(* Asserts that parse rejects header with the expected reason and allocates nothing. *)
METHOD _expectRejected
VAR_INPUT
	header: T_MaxString;
	expected: E_TraceStateFailureReason;
END_VAR
VAR
	_pTraceState: POINTER TO FB_TraceState;
	_success: BOOL;
	_reason: E_TraceStateFailureReason;
END_VAR
_success := TraceStateFactory.parse(pDest:=_pTraceState, pHeader:=ADR(header), failureReason=>_reason);
THIS^.AssertFalse(_success, CONCAT('Expected parse to reject: ', header));
THIS^.AssertEquals_UDINT(TO_UDINT(expected), TO_UDINT(_reason), CONCAT('Expected the failure reason for: ', header));
THIS^.AssertTrue(_pTraceState = 0, CONCAT('Expected nothing to be allocated for: ', header));
IF _pTraceState <> 0 THEN _pTraceState^.delete(pSelf:=_pTraceState); END_IF
END_METHOD

(*
	Writes a valid 515 character header: four 128 character entries k0..k3 joined by ','.
	It is built byte by byte because STRING functions stop at 255 characters.
*)
METHOD _fillLongHeader
VAR_IN_OUT
	header: STRING(600);
END_VAR
VAR
	_p: POINTER TO BYTE;
	_entry: UDINT;
	_i: UDINT;
	_n: UDINT;
END_VAR
_p := ADR(header);
FOR _entry := 0 TO 3 DO
	IF _entry > 0 THEN
		_p[_n] := 16#2C;  // ','
		_n := _n + 1;
	END_IF
	_p[_n] := 16#6B;  // 'k'
	_p[_n + 1] := 16#30 + TO_BYTE(_entry);
	_p[_n + 2] := 16#3D;  // '='
	_n := _n + 3;
	FOR _i := 1 TO 125 DO
		_p[_n] := 16#61 + TO_BYTE(_i MOD 26);
		_n := _n + 1;
	END_FOR
END_FOR
_p[_n] := 0;
END_METHOD

(* parse drops empty members and the optional whitespace around ',' and keeps the order. *)
METHOD testParseCanonicalises : REFERENCE TO FB_Test
VAR
	header: T_MaxString := ' vendor=abc ,, rojo=00f067aa0ba902b7$T, congo@t61rcwkgmze=x ';
	expected: T_MaxString := 'vendor=abc,rojo=00f067aa0ba902b7,congo@t61rcwkgmze=x';
	pTraceState: POINTER TO FB_TraceState;
	success: BOOL;
	reason: E_TraceStateFailureReason;
END_VAR
TcUnit.TEST('testParseCanonicalises');
	success := TraceStateFactory.parse(pDest:=pTraceState, pHeader:=ADR(header), failureReason=>reason);
	THIS^.AssertTrue(success, 'Expected a valid header to parse');
	THIS^.AssertEquals_UDINT(TO_UDINT(E_TraceStateFailureReason.NA), TO_UDINT(reason), 'Expected no failure reason');
	THIS^.AssertTrue(pTraceState <> 0, 'Expected a trace state');
	IF pTraceState <> 0 THEN
		THIS^.AssertEquals_STRING(expected, pTraceState^.pString^, 'Expected the canonical header');
		THIS^.AssertEquals_UDINT(TO_UDINT(LEN(expected)), pTraceState^.length, 'Expected the canonical length');
		THIS^.AssertEquals_UDINT(3, pTraceState^.count, 'Expected three entries');
		pTraceState^.delete(pSelf:=pTraceState);
		THIS^.AssertTrue(pTraceState = 0, 'Expected delete to clear the pointer');
	END_IF
TcUnit.TEST_FINISHED();
END_METHOD

(* An empty header, or one of only empty members, is valid but holds nothing, so no trace state is allocated. *)
METHOD testParseEmptyHeader : REFERENCE TO FB_Test
VAR
	empty: T_MaxString := '';
	blank: T_MaxString := ' , ,,$T';
	pTraceState: POINTER TO FB_TraceState;
	success: BOOL;
	reason: E_TraceStateFailureReason;
END_VAR
TcUnit.TEST('testParseEmptyHeader');
	success := TraceStateFactory.parse(pDest:=pTraceState, pHeader:=ADR(empty), failureReason=>reason);
	THIS^.AssertTrue(success, 'Expected an empty header to be accepted');
	THIS^.AssertEquals_UDINT(TO_UDINT(E_TraceStateFailureReason.NA), TO_UDINT(reason), 'Expected no failure reason');
	THIS^.AssertTrue(pTraceState = 0, 'Expected no trace state for an empty header');

	success := TraceStateFactory.parse(pDest:=pTraceState, pHeader:=ADR(blank), failureReason=>reason);
	THIS^.AssertTrue(success, 'Expected a header of empty members to be accepted');
	THIS^.AssertTrue(pTraceState = 0, 'Expected no trace state for a header of empty members');
	IF pTraceState <> 0 THEN pTraceState^.delete(pSelf:=pTraceState); END_IF
TcUnit.TEST_FINISHED();
END_METHOD

(* Anything that breaks the W3C key or value grammar, or repeats a key, is rejected whole. *)
METHOD testParseRejectsInvalidHeaders : REFERENCE TO FB_Test
VAR
	pTraceState: POINTER TO FB_TraceState;
	pOther: POINTER TO FB_TraceState;
	header: T_MaxString := 'vendor=abc';
	success: BOOL;
	reason: E_TraceStateFailureReason;
END_VAR
TcUnit.TEST('testParseRejectsInvalidHeaders');
	THIS^._expectRejected(header:='Vendor=abc', expected:=E_TraceStateFailureReason.INVALID_KEY);
	THIS^._expectRejected(header:='1vendor=x', expected:=E_TraceStateFailureReason.INVALID_KEY);
	THIS^._expectRejected(header:='=x', expected:=E_TraceStateFailureReason.INVALID_KEY);
	THIS^._expectRejected(header:='@sys=x', expected:=E_TraceStateFailureReason.INVALID_KEY);
	THIS^._expectRejected(header:='tenant@=x', expected:=E_TraceStateFailureReason.INVALID_KEY);
	THIS^._expectRejected(header:='tenant@1sys=x', expected:=E_TraceStateFailureReason.INVALID_KEY);
	THIS^._expectRejected(header:='a@b@c=x', expected:=E_TraceStateFailureReason.INVALID_KEY);
	THIS^._expectRejected(header:='ven dor=x', expected:=E_TraceStateFailureReason.INVALID_KEY);
	THIS^._expectRejected(header:='vendor', expected:=E_TraceStateFailureReason.INVALID_VALUE);
	THIS^._expectRejected(header:='vendor=', expected:=E_TraceStateFailureReason.INVALID_VALUE);
	THIS^._expectRejected(header:='vendor=a=b', expected:=E_TraceStateFailureReason.INVALID_VALUE);
	THIS^._expectRejected(header:='vendor=a$Tb', expected:=E_TraceStateFailureReason.INVALID_VALUE);
	THIS^._expectRejected(header:='good=1,vendor=a=b', expected:=E_TraceStateFailureReason.INVALID_VALUE);
	THIS^._expectRejected(header:='a=1,b=2,a=3', expected:=E_TraceStateFailureReason.DUPLICATE_KEY);

	success := TraceStateFactory.parse(pDest:=pTraceState, pHeader:=0, failureReason=>reason);
	THIS^.AssertFalse(success, 'Expected a null header pointer to be rejected');
	THIS^.AssertEquals_UDINT(TO_UDINT(E_TraceStateFailureReason.HEADER_POINTER_NULL), TO_UDINT(reason), 'Expected HEADER_POINTER_NULL');

	TraceStateFactory.parse(pDest:=pTraceState, pHeader:=ADR(header));
	pOther := pTraceState;
	success := TraceStateFactory.parse(pDest:=pTraceState, pHeader:=ADR(header), failureReason=>reason);
	THIS^.AssertFalse(success, 'Expected an assigned destination to be rejected');
	THIS^.AssertEquals_UDINT(TO_UDINT(E_TraceStateFailureReason.DESTINATION_ALREADY_ASSIGNED), TO_UDINT(reason), 'Expected DESTINATION_ALREADY_ASSIGNED');
	THIS^.AssertTrue(pTraceState = pOther, 'Expected the destination to be left alone');
	IF pTraceState <> 0 THEN pTraceState^.delete(pSelf:=pTraceState); END_IF
TcUnit.TEST_FINISHED();
END_METHOD

(* W3C allows at most 32 entries; a 33rd is rejected. *)
METHOD testParseEntryLimit : REFERENCE TO FB_Test
VAR
	header: T_MaxString;
	i: UDINT;
	pTraceState: POINTER TO FB_TraceState;
	success: BOOL;
	reason: E_TraceStateFailureReason;
END_VAR
TcUnit.TEST('testParseEntryLimit');
	header := 'k0=1';
	FOR i := 1 TO 31 DO
		header := CONCAT(header, CONCAT(CONCAT(',k', UDINT_TO_STRING(i)), '=1'));
	END_FOR
	success := TraceStateFactory.parse(pDest:=pTraceState, pHeader:=ADR(header), failureReason=>reason);
	THIS^.AssertTrue(success, 'Expected 32 entries to be accepted');
	IF pTraceState <> 0 THEN
		THIS^.AssertEquals_UDINT(32, pTraceState^.count, 'Expected 32 entries');
		pTraceState^.delete(pSelf:=pTraceState);
	END_IF

	header := CONCAT(header, ',k32=1');
	success := TraceStateFactory.parse(pDest:=pTraceState, pHeader:=ADR(header), failureReason=>reason);
	THIS^.AssertFalse(success, 'Expected 33 entries to be rejected');
	THIS^.AssertEquals_UDINT(TO_UDINT(E_TraceStateFailureReason.TOO_MANY_ENTRIES), TO_UDINT(reason), 'Expected TOO_MANY_ENTRIES');
	THIS^.AssertTrue(pTraceState = 0, 'Expected nothing to be allocated');
TcUnit.TEST_FINISHED();
END_METHOD

(* A header longer than T_MaxString is kept whole; W3C asks for at least 512 characters. *)
METHOD testParseLongHeader : REFERENCE TO FB_Test
VAR
	header: STRING(600);
	pTraceState: POINTER TO FB_TraceState;
	success: BOOL;
END_VAR
TcUnit.TEST('testParseLongHeader');
	THIS^._fillLongHeader(header:=header);
	THIS^.AssertEquals_UDINT(515, TO_UDINT(LEN2(ADR(header))), 'Expected a 515 character test header');
	success := TraceStateFactory.parse(pDest:=pTraceState, pHeader:=ADR(header));
	THIS^.AssertTrue(success, 'Expected the long header to parse');
	IF pTraceState <> 0 THEN
		THIS^.AssertEquals_UDINT(515, pTraceState^.length, 'Expected all 515 characters');
		THIS^.AssertEquals_UDINT(4, pTraceState^.count, 'Expected four entries');
		THIS^.AssertTrue(MEMCMP(pTraceState^.pString, ADR(header), 516) = 0, 'Expected the header unchanged, with its terminator');
		pTraceState^.delete(pSelf:=pTraceState);
	END_IF
TcUnit.TEST_FINISHED();
END_METHOD

(* clone owns its own buffer, so it outlives the source. *)
METHOD testCloneIsIndependent : REFERENCE TO FB_Test
VAR
	header: T_MaxString := 'vendor=abc,rojo=1';
	pSource: POINTER TO FB_TraceState;
	pClone: POINTER TO FB_TraceState;
	pOther: POINTER TO FB_TraceState;
	success: BOOL;
	reason: E_TraceStateFailureReason;
END_VAR
TcUnit.TEST('testCloneIsIndependent');
	TraceStateFactory.parse(pDest:=pSource, pHeader:=ADR(header));
	success := TraceStateFactory.clone(pDest:=pClone, pSrc:=pSource, failureReason=>reason);
	THIS^.AssertTrue(success, 'Expected clone to succeed');
	THIS^.AssertTrue(pClone <> 0 AND pClone <> pSource, 'Expected a new trace state');
	IF pSource <> 0 AND pClone <> 0 THEN
		THIS^.AssertTrue(pClone^.pString <> pSource^.pString, 'Expected the clone to own its own buffer');
	END_IF

	success := TraceStateFactory.clone(pDest:=pClone, pSrc:=pSource, failureReason=>reason);
	THIS^.AssertFalse(success, 'Expected clone into an assigned destination to fail');
	THIS^.AssertEquals_UDINT(TO_UDINT(E_TraceStateFailureReason.DESTINATION_ALREADY_ASSIGNED), TO_UDINT(reason), 'Expected DESTINATION_ALREADY_ASSIGNED');
	success := TraceStateFactory.clone(pDest:=pOther, pSrc:=0, failureReason=>reason);
	THIS^.AssertFalse(success, 'Expected clone of a null source to fail');
	THIS^.AssertEquals_UDINT(TO_UDINT(E_TraceStateFailureReason.SOURCE_POINTER_NULL), TO_UDINT(reason), 'Expected SOURCE_POINTER_NULL');

	IF pSource <> 0 THEN pSource^.delete(pSelf:=pSource); END_IF
	IF pClone <> 0 THEN
		THIS^.AssertEquals_STRING('vendor=abc,rojo=1', pClone^.pString^, 'Expected the clone to outlive its source');
		THIS^.AssertEquals_UDINT(2, pClone^.count, 'Expected the entry count to be copied');
		pClone^.delete(pSelf:=pClone);
	END_IF
TcUnit.TEST_FINISHED();
END_METHOD

(* truncate removes entries over 128 characters first, then entries from the right, and never cuts an entry. *)
METHOD testTruncateFollowsW3C : REFERENCE TO FB_Test
VAR
	header: STRING(600);
	pBytes: POINTER TO BYTE;
	i: UDINT;
	pSource: POINTER TO FB_TraceState;
	pResult: POINTER TO FB_TraceState;
	success: BOOL;
	reason: E_TraceStateFailureReason;
END_VAR
TcUnit.TEST('testTruncateFollowsW3C');
	// a=1,big=<130 characters>,b=2,c=3
	header := 'a=1,big=';
	pBytes := ADR(header);
	FOR i := 8 TO 137 DO
		pBytes[i] := 16#78;  // 'x'
	END_FOR
	pBytes[138] := 0;
	MEMCPY(pBytes + 138, ADR(',b=2,c=3'), 9);
	success := TraceStateFactory.parse(pDest:=pSource, pHeader:=ADR(header));
	THIS^.AssertTrue(success AND pSource <> 0, 'Expected the header to parse');
	IF pSource = 0 THEN
		TcUnit.TEST_FINISHED();
		RETURN;
	END_IF
	THIS^.AssertEquals_UDINT(146, pSource^.length, 'Expected a 146 character test header');

	success := TraceStateFactory.truncate(pDest:=pResult, pSrc:=pSource, maxLength:=1000, failureReason=>reason);
	THIS^.AssertTrue(success AND pResult <> 0, 'Expected a header that fits to be copied');
	IF pResult <> 0 THEN
		THIS^.AssertTrue(pResult <> pSource AND pResult^.length = 146, 'Expected a whole copy');
		pResult^.delete(pSelf:=pResult);
	END_IF

	success := TraceStateFactory.truncate(pDest:=pResult, pSrc:=pSource, maxLength:=20, failureReason=>reason);
	THIS^.AssertTrue(success, 'Expected truncate to succeed');
	IF pResult <> 0 THEN
		THIS^.AssertEquals_STRING('a=1,b=2,c=3', pResult^.pString^, 'Expected the large entry to go first');
		THIS^.AssertEquals_UDINT(3, pResult^.count, 'Expected three entries');
		pResult^.delete(pSelf:=pResult);
	ELSE
		THIS^.AssertTrue(FALSE, 'Expected a truncated trace state');
	END_IF

	success := TraceStateFactory.truncate(pDest:=pResult, pSrc:=pSource, maxLength:=7, failureReason=>reason);
	THIS^.AssertTrue(success, 'Expected truncate to succeed');
	IF pResult <> 0 THEN
		THIS^.AssertEquals_STRING('a=1,b=2', pResult^.pString^, 'Expected entries to go from the right next');
		pResult^.delete(pSelf:=pResult);
	ELSE
		THIS^.AssertTrue(FALSE, 'Expected a truncated trace state');
	END_IF

	success := TraceStateFactory.truncate(pDest:=pResult, pSrc:=pSource, maxLength:=2, failureReason=>reason);
	THIS^.AssertTrue(success, 'Expected truncate to succeed when nothing fits');
	THIS^.AssertTrue(pResult = 0, 'Expected no trace state when no entry fits');
	IF pResult <> 0 THEN pResult^.delete(pSelf:=pResult); END_IF

	success := TraceStateFactory.truncate(pDest:=pResult, pSrc:=0, maxLength:=512, failureReason=>reason);
	THIS^.AssertFalse(success, 'Expected a null source to be rejected');
	THIS^.AssertEquals_UDINT(TO_UDINT(E_TraceStateFailureReason.SOURCE_POINTER_NULL), TO_UDINT(reason), 'Expected SOURCE_POINTER_NULL');

	pSource^.delete(pSelf:=pSource);
TcUnit.TEST_FINISHED();
END_METHOD

END_FUNCTION_BLOCK

// ---- TEST/TRACING/PROPAGATION/FB_TestTraceContextPropagator.TcPOU
(* Tests TraceContextPropagator.extract and inject against the W3C traceparent and tracestate rules. *)
FUNCTION_BLOCK FB_TestTraceContextPropagator EXTENDS FB_TestSuite

THIS^.testExtractsTraceparentAndTracestate();
THIS^.testKeepsUnsampledFlag();
THIS^.testAcceptsFutureVersion();
THIS^.testMeasuresTraceparentBeyond255();
THIS^.testTracestateIsOptional();
THIS^.testKeepsLongTracestateWhole();
THIS^.testRejectsMalformedTraceparent();
THIS^.testRejectsAssignedDestination();
THIS^.testInjectWritesExtractedCarrier();
THIS^.testInjectDropsWholeTracestateEntries();
THIS^.testInjectRejectsMissingOrInvalidContext();

(*
	Asserts that extract rejects traceparent with the expected reason and leaves the destination
	at 0. The tracestate beside it is valid, so this also shows a bad traceparent drops it.
*)
METHOD _expectRejected
VAR_INPUT
	traceparent: T_MaxString;  // longer than 55, so overlong headers reach extract whole
	expected: E_PropagationFailureReason;
END_VAR
VAR
	_pContext: POINTER TO FB_SpanContext;
	_success: BOOL;
	_reason: E_PropagationFailureReason;
END_VAR
_success := TraceContextPropagator.extract(
	pDest:=_pContext,
	traceparent:=traceparent,
	tracestate:='vendor=abc',
	failureReason=>_reason
);
THIS^.AssertFalse(_success, CONCAT('Expected extract to reject: ', traceparent));
THIS^.AssertEquals_UDINT(TO_UDINT(expected), TO_UDINT(_reason), CONCAT('Expected the failure reason for: ', traceparent));
THIS^.AssertTrue(_pContext = 0, CONCAT('Expected no context for: ', traceparent));
IF _pContext <> 0 THEN _pContext^.delete(pSelf:=_pContext); END_IF
END_METHOD

(*
	The W3C example carrier becomes a remote context holding the caller's trace id, span id,
	sampled bit and tracestate, so a PLC span can link back to the span that triggered it.
*)
METHOD testExtractsTraceparentAndTracestate : REFERENCE TO FB_Test
VAR
	traceparent: STRING(55) := '00-4bf92f3577b34da6a3ce929d0e0e4736-00f067aa0ba902b7-01';
	tracestate: STRING(512) := 'congo=t61rcWkgMzE,rojo=00f067aa0ba902b7';
	expectedTraceId: ARRAY [0..15] OF BYTE := [
		16#4B, 16#F9, 16#2F, 16#35, 16#77, 16#B3, 16#4D, 16#A6,
		16#A3, 16#CE, 16#92, 16#9D, 16#0E, 16#0E, 16#47, 16#36];
	expectedSpanId: ARRAY [0..7] OF BYTE := [16#00, 16#F0, 16#67, 16#AA, 16#0B, 16#A9, 16#02, 16#B7];
	pContext: POINTER TO FB_SpanContext;
	pTraceState: POINTER TO FB_TraceState;
	traceId: REFERENCE TO FB_TraceId;
	spanId: REFERENCE TO FB_SpanId;
	success: BOOL;
	reason: E_PropagationFailureReason;
END_VAR
TcUnit.TEST('testExtractsTraceparentAndTracestate');
	success := TraceContextPropagator.extract(
		pDest:=pContext,
		traceparent:=traceparent,
		tracestate:=tracestate,
		failureReason=>reason
	);
	THIS^.AssertTrue(success, 'Expected the W3C example carrier to be extracted');
	THIS^.AssertEquals_UDINT(TO_UDINT(E_PropagationFailureReason.NA), TO_UDINT(reason), 'Expected no failure reason on success');
	THIS^.AssertTrue(pContext <> 0, 'Expected extract to assign the destination');
	IF pContext = 0 THEN
		TcUnit.TEST_FINISHED();
		RETURN;
	END_IF

	traceId REF= pContext^.traceId;
	spanId REF= pContext^.spanId;
	THIS^.AssertTrue(
		MEMCMP(ADR(traceId.bytes), ADR(expectedTraceId), SIZEOF(expectedTraceId)) = 0,
		'Expected the trace id decoded from the traceparent'
	);
	THIS^.AssertTrue(
		MEMCMP(ADR(spanId.bytes), ADR(expectedSpanId), SIZEOF(expectedSpanId)) = 0,
		'Expected the caller$'s span id decoded from the traceparent'
	);
	THIS^.AssertEquals_UDINT(16#301, pContext^.traceFlags, 'Expected the sampled bit and both remote bits');
	THIS^.AssertTrue(pContext^.isRemote(), 'Expected an extracted context to be remote');

	pTraceState := pContext^.traceState;
	THIS^.AssertTrue(pTraceState <> 0, 'Expected the tracestate to be kept');
	IF pTraceState <> 0 THEN
		THIS^.AssertEquals_STRING('congo=t61rcWkgMzE,rojo=00f067aa0ba902b7', pTraceState^.pString^, 'Expected the tracestate entries in their original order');
	END_IF
	pContext^.delete(pSelf:=pContext);
TcUnit.TEST_FINISHED();
END_METHOD

(*
	A caller that did not sample its own trace still produces a context: the sampled bit is
	carried as sent, and the default sampler does not sample a child of the context.
*)
METHOD testKeepsUnsampledFlag : REFERENCE TO FB_Test
VAR
	traceparent: STRING(55) := '00-4bf92f3577b34da6a3ce929d0e0e4736-00f067aa0ba902b7-00';
	pContext: POINTER TO FB_SpanContext;
	success: BOOL;
END_VAR
TcUnit.TEST('testKeepsUnsampledFlag');
	success := TraceContextPropagator.extract(pDest:=pContext, traceparent:=traceparent, tracestate:='');
	THIS^.AssertTrue(success, 'Expected an unsampled carrier to be extracted');
	IF pContext <> 0 THEN
		THIS^.AssertEquals_UDINT(16#300, pContext^.traceFlags, 'Expected both remote bits and no sampled bit');
		THIS^.AssertTrue(pContext^.isRemote(), 'Expected an extracted context to be remote');
		pContext^.delete(pSelf:=pContext);
	END_IF
TcUnit.TEST_FINISHED();
END_METHOD

(*
	W3C asks a parser to read a newer version as version 00 rather than reject it, ignoring any
	fields after the flags, so a caller that upgrades its tracing library does not lose the link.
	The flags may end the header or be followed by '-' and more fields.
*)
METHOD testAcceptsFutureVersion : REFERENCE TO FB_Test
VAR
	traceparent: STRING(80) := 'cc-4bf92f3577b34da6a3ce929d0e0e4736-00f067aa0ba902b7-01-newfield';
	traceparentWithoutFields: STRING(55) := 'cc-4bf92f3577b34da6a3ce929d0e0e4736-00f067aa0ba902b7-01';
	pContext: POINTER TO FB_SpanContext;
	success: BOOL;
	reason: E_PropagationFailureReason;
END_VAR
TcUnit.TEST('testAcceptsFutureVersion');
	success := TraceContextPropagator.extract(pDest:=pContext, traceparent:=traceparent, tracestate:='', failureReason=>reason);
	THIS^.AssertTrue(success, 'Expected version cc with an extra field to be read as version 00');
	THIS^.AssertEquals_UDINT(TO_UDINT(E_PropagationFailureReason.NA), TO_UDINT(reason), 'Expected no failure reason for a future version');
	IF pContext <> 0 THEN pContext^.delete(pSelf:=pContext); END_IF

	// the flags end the header
	success := TraceContextPropagator.extract(pDest:=pContext, traceparent:=traceparentWithoutFields, tracestate:='', failureReason=>reason);
	THIS^.AssertTrue(success, 'Expected version cc with no extra field to be read as version 00');
	THIS^.AssertEquals_UDINT(TO_UDINT(E_PropagationFailureReason.NA), TO_UDINT(reason), 'Expected no failure reason for a 55 character future version');
	IF pContext <> 0 THEN pContext^.delete(pSelf:=pContext); END_IF
TcUnit.TEST_FINISHED();
END_METHOD

(*
	The traceparent alone identifies the caller's span. A missing tracestate, or one that breaks
	the W3C grammar, leaves the context without a trace state instead of failing the extraction.
*)
METHOD testTracestateIsOptional : REFERENCE TO FB_Test
VAR
	traceparent: STRING(55) := '00-4bf92f3577b34da6a3ce929d0e0e4736-00f067aa0ba902b7-01';
	pContext: POINTER TO FB_SpanContext;
	success: BOOL;
	reason: E_PropagationFailureReason;
END_VAR
TcUnit.TEST('testTracestateIsOptional');
	// no tracestate header
	success := TraceContextPropagator.extract(pDest:=pContext, traceparent:=traceparent, tracestate:='', failureReason=>reason);
	THIS^.AssertTrue(success, 'Expected a carrier without tracestate to be extracted');
	THIS^.AssertTrue(pContext <> 0 AND_THEN pContext^.traceState = 0, 'Expected no trace state without a tracestate header');
	IF pContext <> 0 THEN pContext^.delete(pSelf:=pContext); END_IF

	// an uppercase key breaks the tracestate grammar, so only the trace state is dropped
	success := TraceContextPropagator.extract(pDest:=pContext, traceparent:=traceparent, tracestate:='Vendor=abc', failureReason=>reason);
	THIS^.AssertTrue(success, 'Expected an invalid tracestate not to fail the extraction');
	THIS^.AssertEquals_UDINT(TO_UDINT(E_PropagationFailureReason.NA), TO_UDINT(reason), 'Expected no failure reason for a dropped tracestate');
	THIS^.AssertTrue(pContext <> 0 AND_THEN pContext^.traceState = 0, 'Expected an invalid tracestate to be dropped');
	IF pContext <> 0 THEN pContext^.delete(pSelf:=pContext); END_IF
TcUnit.TEST_FINISHED();
END_METHOD

(*
	Each way a traceparent can break the W3C format is reported by its own reason, and nothing
	is allocated, so the caller can start an unlinked span and log why.
*)
METHOD testRejectsMalformedTraceparent : REFERENCE TO FB_Test
TcUnit.TEST('testRejectsMalformedTraceparent');
	// no header at all
	THIS^._expectRejected(traceparent:='', expected:=E_PropagationFailureReason.TRACEPARENT_EMPTY);
	// the flags are missing
	THIS^._expectRejected(traceparent:='00-4bf92f3577b34da6a3ce929d0e0e4736-00f067aa0ba902b7', expected:=E_PropagationFailureReason.TRACEPARENT_LENGTH_INVALID);
	// version ff is reserved as invalid
	THIS^._expectRejected(traceparent:='ff-4bf92f3577b34da6a3ce929d0e0e4736-00f067aa0ba902b7-01', expected:=E_PropagationFailureReason.VERSION_INVALID);
	// the version is not hex
	THIS^._expectRejected(traceparent:='0g-4bf92f3577b34da6a3ce929d0e0e4736-00f067aa0ba902b7-01', expected:=E_PropagationFailureReason.VERSION_INVALID);
	// the version is not followed by '-'
	THIS^._expectRejected(traceparent:='00_4bf92f3577b34da6a3ce929d0e0e4736-00f067aa0ba902b7-01', expected:=E_PropagationFailureReason.DELIMITER_INVALID);
	// W3C allows only lowercase hex
	THIS^._expectRejected(traceparent:='00-4BF92F3577B34DA6A3CE929D0E0E4736-00f067aa0ba902b7-01', expected:=E_PropagationFailureReason.TRACE_ID_INVALID);
	// an all-zero trace id means absent
	THIS^._expectRejected(traceparent:='00-00000000000000000000000000000000-00f067aa0ba902b7-01', expected:=E_PropagationFailureReason.TRACE_ID_INVALID);
	// the span id is not hex
	THIS^._expectRejected(traceparent:='00-4bf92f3577b34da6a3ce929d0e0e4736-00f067aa0ba902bx-01', expected:=E_PropagationFailureReason.SPAN_ID_INVALID);
	// an all-zero span id means absent
	THIS^._expectRejected(traceparent:='00-4bf92f3577b34da6a3ce929d0e0e4736-0000000000000000-01', expected:=E_PropagationFailureReason.SPAN_ID_INVALID);
	// the flags are not hex
	THIS^._expectRejected(traceparent:='00-4bf92f3577b34da6a3ce929d0e0e4736-00f067aa0ba902b7-0z', expected:=E_PropagationFailureReason.TRACE_FLAGS_INVALID);
	// version 00 is exactly 55 characters, so nothing may follow the flags
	THIS^._expectRejected(traceparent:='00-4bf92f3577b34da6a3ce929d0e0e4736-00f067aa0ba902b7-01-00', expected:=E_PropagationFailureReason.TRACEPARENT_LENGTH_INVALID);
	// a future version's flags must be followed by '-' or the end of the header
	THIS^._expectRejected(traceparent:='cc-4bf92f3577b34da6a3ce929d0e0e4736-00f067aa0ba902b7-01x', expected:=E_PropagationFailureReason.DELIMITER_INVALID);
TcUnit.TEST_FINISHED();
END_METHOD

(* extract never overwrites a context the caller already owns, which would leak it. *)
METHOD testRejectsAssignedDestination : REFERENCE TO FB_Test
VAR
	traceparent: STRING(55) := '00-4bf92f3577b34da6a3ce929d0e0e4736-00f067aa0ba902b7-01';
	pContext: POINTER TO FB_SpanContext;
	pFirst: POINTER TO FB_SpanContext;
	success: BOOL;
	reason: E_PropagationFailureReason;
END_VAR
TcUnit.TEST('testRejectsAssignedDestination');
	TraceContextPropagator.extract(pDest:=pContext, traceparent:=traceparent, tracestate:='');
	pFirst := pContext;

	success := TraceContextPropagator.extract(pDest:=pContext, traceparent:=traceparent, tracestate:='', failureReason=>reason);
	THIS^.AssertFalse(success, 'Expected extract to refuse an assigned destination');
	THIS^.AssertEquals_UDINT(
		TO_UDINT(E_PropagationFailureReason.DESTINATION_ALREADY_ASSIGNED),
		TO_UDINT(reason),
		'Expected DESTINATION_ALREADY_ASSIGNED'
	);
	THIS^.AssertTrue(pContext = pFirst, 'Expected the caller$'s context to be left in place');
	IF pContext <> 0 THEN pContext^.delete(pSelf:=pContext); END_IF
TcUnit.TEST_FINISHED();
END_METHOD

(*
	Writes a valid 515 character tracestate: four 128 character entries k0..k3 joined by ','.
	It is built byte by byte because STRING functions stop at 255 characters.
*)
METHOD _fillLongHeader
VAR_IN_OUT
	header: STRING(600);
END_VAR
VAR
	_p: POINTER TO BYTE;
	_entry: UDINT;
	_i: UDINT;
	_n: UDINT;
END_VAR
_p := ADR(header);
FOR _entry := 0 TO 3 DO
	IF _entry > 0 THEN
		_p[_n] := 16#2C;  // ','
		_n := _n + 1;
	END_IF
	_p[_n] := 16#6B;  // 'k'
	_p[_n + 1] := 16#30 + TO_BYTE(_entry);
	_p[_n + 2] := 16#3D;  // '='
	_n := _n + 3;
	FOR _i := 1 TO 125 DO
		_p[_n] := 16#61 + TO_BYTE(_i MOD 26);
		_n := _n + 1;
	END_FOR
END_FOR
_p[_n] := 0;
END_METHOD

(*
	W3C asks for at least 512 tracestate characters to be kept and allows dropping only whole
	entries, never cutting one. A 515 character header is kept entirely, so no vendor's entry
	reaches the backend corrupted.
*)
METHOD testKeepsLongTracestateWhole : REFERENCE TO FB_Test
VAR
	traceparent: STRING(55) := '00-4bf92f3577b34da6a3ce929d0e0e4736-00f067aa0ba902b7-01';
	tracestate: STRING(600);
	pContext: POINTER TO FB_SpanContext;
	pTraceState: POINTER TO FB_TraceState;
	success: BOOL;
END_VAR
TcUnit.TEST('testKeepsLongTracestateWhole');
	THIS^._fillLongHeader(header:=tracestate);
	success := TraceContextPropagator.extract(pDest:=pContext, traceparent:=traceparent, tracestate:=tracestate);
	THIS^.AssertTrue(success, 'Expected a carrier with a long tracestate to be extracted');
	IF pContext <> 0 THEN
		pTraceState := pContext^.traceState;
		THIS^.AssertTrue(pTraceState <> 0, 'Expected the long tracestate to be kept');
		IF pTraceState <> 0 THEN
			THIS^.AssertEquals_UDINT(515, pTraceState^.length, 'Expected all 515 characters, with no entry cut');
			THIS^.AssertEquals_UDINT(4, pTraceState^.count, 'Expected all four entries');
		END_IF
		pContext^.delete(pSelf:=pContext);
	END_IF
TcUnit.TEST_FINISHED();
END_METHOD

(*
	A carrier can be longer than the 255 characters that LEN and T_MaxString handle. extract
	measures the whole header, so a 300 character version 00 header is still rejected and a
	300 character future version with extra fields is still accepted.
*)
METHOD testMeasuresTraceparentBeyond255 : REFERENCE TO FB_Test
VAR
	versionZero: STRING(300);
	futureVersion: STRING(300);
	pContext: POINTER TO FB_SpanContext;
	success: BOOL;
	reason: E_PropagationFailureReason;
END_VAR
TcUnit.TEST('testMeasuresTraceparentBeyond255');
	THIS^._fillLongTraceparent(header:=versionZero, prefix:='00-4bf92f3577b34da6a3ce929d0e0e4736-00f067aa0ba902b7-01');
	THIS^._fillLongTraceparent(header:=futureVersion, prefix:='cc-4bf92f3577b34da6a3ce929d0e0e4736-00f067aa0ba902b7-01');

	success := TraceContextPropagator.extract(pDest:=pContext, traceparent:=versionZero, tracestate:='', failureReason=>reason);
	THIS^.AssertFalse(success, 'Expected a 300 character version 00 traceparent to be rejected');
	THIS^.AssertEquals_UDINT(TO_UDINT(E_PropagationFailureReason.TRACEPARENT_LENGTH_INVALID), TO_UDINT(reason), 'Expected TRACEPARENT_LENGTH_INVALID for a 300 character version 00 traceparent');
	THIS^.AssertTrue(pContext = 0, 'Expected no context for a 300 character version 00 traceparent');
	IF pContext <> 0 THEN pContext^.delete(pSelf:=pContext); END_IF

	success := TraceContextPropagator.extract(pDest:=pContext, traceparent:=futureVersion, tracestate:='', failureReason=>reason);
	THIS^.AssertTrue(success, 'Expected a 300 character future version traceparent to be accepted');
	THIS^.AssertEquals_UDINT(TO_UDINT(E_PropagationFailureReason.NA), TO_UDINT(reason), 'Expected no failure reason for a 300 character future version traceparent');
	IF pContext <> 0 THEN pContext^.delete(pSelf:=pContext); END_IF
TcUnit.TEST_FINISHED();
END_METHOD

(*
	Writes a 300 character traceparent: the 55 character prefix, then '-' and 244 'a' characters
	as extra fields. It is built byte by byte because STRING functions stop at 255 characters.
*)
METHOD _fillLongTraceparent
VAR_IN_OUT
	header: STRING(300);
END_VAR
VAR_INPUT
	prefix: STRING(55);
END_VAR
VAR
	_p: POINTER TO BYTE;
	_i: UDINT;
END_VAR
header := prefix;
_p := ADR(header);
_p[55] := 16#2D;  // '-'
FOR _i := 56 TO 299 DO
	_p[_i] := 16#61;  // 'a'
END_FOR
_p[300] := 0;
END_METHOD

(*
	inject is the inverse of extract: a context extracted from the W3C example carrier writes the
	same traceparent and tracestate back out, so a context forwarded by the PLC reaches the next
	service unchanged. The remote bits stay behind, because they are OTLP flags, not W3C flags.
*)
METHOD testInjectWritesExtractedCarrier : REFERENCE TO FB_Test
VAR
	traceparentIn: STRING(55) := '00-4bf92f3577b34da6a3ce929d0e0e4736-00f067aa0ba902b7-01';
	tracestateIn: STRING(512) := 'congo=t61rcWkgMzE,rojo=00f067aa0ba902b7';
	carrier: ST_TraceContextCarrier;
	pContext: POINTER TO FB_SpanContext;
	success: BOOL;
	reason: E_PropagationFailureReason;
END_VAR
TcUnit.TEST('testInjectWritesExtractedCarrier');
	TraceContextPropagator.extract(pDest:=pContext, traceparent:=traceparentIn, tracestate:=tracestateIn);
	success := TraceContextPropagator.inject(pContext:=pContext, carrier:=carrier, failureReason=>reason);
	THIS^.AssertTrue(success, 'Expected a valid context to be injected');
	THIS^.AssertEquals_UDINT(TO_UDINT(E_PropagationFailureReason.NA), TO_UDINT(reason), 'Expected no failure reason for a valid context');
	THIS^.AssertEquals_STRING(traceparentIn, carrier.traceparent, 'Expected the traceparent that was extracted');
	THIS^.AssertEquals_STRING(tracestateIn, carrier.tracestate, 'Expected the tracestate that was extracted');
	IF pContext <> 0 THEN pContext^.delete(pSelf:=pContext); END_IF
TcUnit.TEST_FINISHED();
END_METHOD

(*
	The inject carrier holds 512 characters, the W3C floor. A longer trace state is shortened by
	dropping whole entries from the right, never by cutting one, so every vendor entry that is
	sent on is still intact.
*)
METHOD testInjectDropsWholeTracestateEntries : REFERENCE TO FB_Test
VAR
	traceparentIn: STRING(55) := '00-4bf92f3577b34da6a3ce929d0e0e4736-00f067aa0ba902b7-01';
	tracestateIn: STRING(600);
	carrier: ST_TraceContextCarrier;
	pContext: POINTER TO FB_SpanContext;
	success: BOOL;
END_VAR
TcUnit.TEST('testInjectDropsWholeTracestateEntries');
	// four 128 character entries k0..k3: 515 characters
	THIS^._fillLongHeader(header:=tracestateIn);
	TraceContextPropagator.extract(pDest:=pContext, traceparent:=traceparentIn, tracestate:=tracestateIn);
	success := TraceContextPropagator.inject(pContext:=pContext, carrier:=carrier);
	THIS^.AssertTrue(success, 'Expected a context with a long trace state to be injected');
	// three whole entries and two commas: 3 * 128 + 2
	THIS^.AssertEquals_UDINT(386, TO_UDINT(LEN2(ADR(carrier.tracestate))), 'Expected k3 to be dropped whole, leaving 386 characters');
	THIS^.AssertTrue(MEMCMP(ADR(carrier.tracestate), ADR(tracestateIn), 386) = 0, 'Expected the first three entries unchanged');
	IF pContext <> 0 THEN pContext^.delete(pSelf:=pContext); END_IF
TcUnit.TEST_FINISHED();
END_METHOD

(*
	There is nothing to propagate without a valid identity. inject fails and leaves both headers
	empty, so the caller sends no header rather than a malformed one.
*)
METHOD testInjectRejectsMissingOrInvalidContext : REFERENCE TO FB_Test
VAR
	traceId: FB_TraceId;  // all zero: the encoding of "absent"
	spanId: FB_SpanId;
	carrier: ST_TraceContextCarrier := (traceparent:='stale', tracestate:='stale=1');
	pContext: POINTER TO FB_SpanContext;
	success: BOOL;
	reason: E_PropagationFailureReason;
END_VAR
TcUnit.TEST('testInjectRejectsMissingOrInvalidContext');
	success := TraceContextPropagator.inject(pContext:=0, carrier:=carrier, failureReason=>reason);
	THIS^.AssertFalse(success, 'Expected inject to reject a null context');
	THIS^.AssertEquals_UDINT(TO_UDINT(E_PropagationFailureReason.CONTEXT_POINTER_NULL), TO_UDINT(reason), 'Expected CONTEXT_POINTER_NULL for a null context');
	THIS^.AssertEquals_STRING('', carrier.traceparent, 'Expected an empty traceparent after a null context');
	THIS^.AssertEquals_STRING('', carrier.tracestate, 'Expected an empty tracestate after a null context');

	// ContextFactory does not validate identities, so it can build the invalid context
	ContextFactory.buildContext(pDest:=pContext, pTraceId:=ADR(traceId), pSpanId:=ADR(spanId), pTraceState:=0, traceFlags:=1);
	success := TraceContextPropagator.inject(pContext:=pContext, carrier:=carrier, failureReason=>reason);
	THIS^.AssertFalse(success, 'Expected inject to reject a context with all-zero ids');
	THIS^.AssertEquals_UDINT(TO_UDINT(E_PropagationFailureReason.CONTEXT_INVALID), TO_UDINT(reason), 'Expected CONTEXT_INVALID for all-zero ids');
	THIS^.AssertEquals_STRING('', carrier.traceparent, 'Expected an empty traceparent after an invalid context');
	IF pContext <> 0 THEN pContext^.delete(pSelf:=pContext); END_IF
TcUnit.TEST_FINISHED();
END_METHOD

END_FUNCTION_BLOCK

// ---- TEST/TRACING/PROPAGATION/FB_TestAdsLoopbackPropagation.TcPOU
(*
	Sends a span context to this PLC over ADS and extracts it on arrival, the way an upstream
	gateway would deliver a carrier. It proves inject, an ADS transport and extract agree end to
	end, and shows that ST_TraceContextCarrier can travel as one ADS write. The test writes to its own _received symbol through a handle on this PLC's ADS port.
*)
FUNCTION_BLOCK FB_TestAdsLoopbackPropagation EXTENDS FB_TestSuite
VAR CONSTANT
	ADSIGRP_SYM_HNDBYNAME: UDINT := 16#F003;  // get a handle for a symbol name
	ADSIGRP_SYM_VALBYHND: UDINT := 16#F005;  // read or write a symbol through its handle
	ADSIGRP_SYM_RELEASEHND: UDINT := 16#F006;  // release a handle
	ADS_TIMEOUT: TIME := T#2S;  // each ADS request gives up after this, so every wait below is bounded
	EXCHANGE_TIMEOUT: TIME := T#5S;  // longer than ADS_TIMEOUT, so an ADS request in flight can still finish
END_VAR
VAR
	// the MAIN instance path of this suite; change it if the instance is renamed
	_symbol: T_MaxString := 'MAIN.fbTestAdsLoopbackPropagation._received';
	_sent: ST_TraceContextCarrier;
	_received: ST_TraceContextCarrier;
	_handle: UDINT;
	_hasHandle: BOOL;
	_getHandle: ADSRDWRT;
	_write: ADSWRITE;
	_releaseHandle: ADSWRITE;
	_state: USINT;
	_exchangeTimer: TON;
	_timedOut: BOOL;  // no new request starts once set; requests in flight still finish
END_VAR

THIS^.testCarrierSurvivesAdsLoopback();

(*
	A context injected into a carrier, written to this PLC over ADS and extracted on arrival has
	the same ids, sampled bit and trace state, and is marked remote. This is the path a gateway
	command takes, so a mismatch here would split the caller's trace from the PLC's.
*)
METHOD testCarrierSurvivesAdsLoopback : REFERENCE TO FB_Test
VAR
	source: STRING(55) := '00-4bf92f3577b34da6a3ce929d0e0e4736-00f067aa0ba902b7-01';
	sourceState: STRING(512) := 'congo=t61rcWkgMzE,rojo=00f067aa0ba902b7';
	pSent: POINTER TO FB_SpanContext;
	pReceived: POINTER TO FB_SpanContext;
	reason: E_PropagationFailureReason;
	pTraceState: POINTER TO FB_TraceState;
END_VAR
TcUnit.TEST('testCarrierSurvivesAdsLoopback');
	// the timeout never abandons a request in flight: each state still waits for its ADS block,
	// which gives up after ADS_TIMEOUT, and then releases the handle if one was granted
	_exchangeTimer(IN:=_state > 0 AND _state < 50, PT:=EXCHANGE_TIMEOUT);
	IF _exchangeTimer.Q AND NOT _timedOut THEN
		THIS^.AssertTrue(FALSE, 'Expected the ADS loopback to finish within EXCHANGE_TIMEOUT');
		_timedOut := TRUE;
	END_IF

	CASE _state OF
		0: // the source context comes from the W3C example carrier; inject writes it back out
			IF NOT TraceContextPropagator.extract(pDest:=pSent, traceparent:=source, tracestate:=sourceState) THEN
				THIS^.AssertTrue(FALSE, 'Expected the source carrier to extract');
				_state := 50;
				RETURN;
			END_IF
			TraceContextPropagator.inject(pContext:=pSent, carrier:=_sent, failureReason=>reason);
			pSent^.delete(pSelf:=pSent);
			THIS^.AssertEquals_UDINT(TO_UDINT(E_PropagationFailureReason.NA), TO_UDINT(reason), 'Expected the source context to inject');
			MEMSET(ADR(_received), 0, SIZEOF(_received));
			// NETID '' is this machine; the port is this PLC's own ADS port
			_getHandle(
				NETID:='',
				PORT:=TwinCAT_SystemInfoVarList._AppInfo.AdsPort,
				IDXGRP:=ADSIGRP_SYM_HNDBYNAME,
				IDXOFFS:=0,
				WRITELEN:=TO_UDINT(LEN(_symbol)),
				READLEN:=SIZEOF(_handle),
				SRCADDR:=ADR(_symbol),
				DESTADDR:=ADR(_handle),
				WRTRD:=TRUE,
				TMOUT:=ADS_TIMEOUT);
			_state := 10;

		10: // wait for the symbol handle
			_getHandle(WRTRD:=FALSE);
			IF NOT _getHandle.BUSY THEN
				IF _getHandle.ERR THEN
					THIS^.AssertTrue(FALSE, CONCAT('Expected a handle for _received, ADS error ', UDINT_TO_STRING(_getHandle.ERRID)));
					_state := 50;
				ELSIF _timedOut THEN
					_hasHandle := TRUE;  // granted late: skip the write, but still release it
					_state := 40;
				ELSE
					_hasHandle := TRUE;
					// both headers in one write, as a gateway's single method call would deliver them
					_write(
						NETID:='',
						PORT:=TwinCAT_SystemInfoVarList._AppInfo.AdsPort,
						IDXGRP:=ADSIGRP_SYM_VALBYHND,
						IDXOFFS:=_handle,
						LEN:=SIZEOF(_sent),
						SRCADDR:=ADR(_sent),
						WRITE:=TRUE,
						TMOUT:=ADS_TIMEOUT);
					_state := 20;
				END_IF
			END_IF

		20: // wait for the write, then extract what arrived
			_write(WRITE:=FALSE);
			IF NOT _write.BUSY THEN
				IF _write.ERR THEN
					THIS^.AssertTrue(FALSE, CONCAT('Expected the carrier write to succeed, ADS error ', UDINT_TO_STRING(_write.ERRID)));
				ELSE
					THIS^.AssertEquals_STRING(_sent.traceparent, _received.traceparent, 'Expected the traceparent to arrive unchanged');
					THIS^.AssertEquals_STRING(_sent.tracestate, _received.tracestate, 'Expected the tracestate to arrive unchanged');
					IF TraceContextPropagator.extract(pDest:=pReceived, traceparent:=_received.traceparent, tracestate:=_received.tracestate, failureReason=>reason) THEN
						// 16#301: sampled, remoteness known, remote
						THIS^.AssertEquals_UDINT(16#301, pReceived^.traceFlags, 'Expected the sampled bit and both remote bits on arrival');
						THIS^.AssertEquals_STRING(source, _received.traceparent, 'Expected the ids and flags of the source carrier');
						pTraceState := pReceived^.traceState;
						THIS^.AssertTrue(pTraceState <> 0, 'Expected the trace state to arrive');
						IF pTraceState <> 0 THEN
							THIS^.AssertEquals_UDINT(2, pTraceState^.count, 'Expected both trace state entries to arrive');
						END_IF
						pReceived^.delete(pSelf:=pReceived);
					ELSE
						THIS^.AssertTrue(FALSE, CONCAT('Expected the received carrier to extract, reason ', TO_STRING(reason)));
					END_IF
				END_IF
				_state := 40;
			END_IF

		40: // release the handle whether or not the exchange succeeded
			IF _hasHandle THEN
				_releaseHandle(
					NETID:='',
					PORT:=TwinCAT_SystemInfoVarList._AppInfo.AdsPort,
					IDXGRP:=ADSIGRP_SYM_RELEASEHND,
					IDXOFFS:=0,
					LEN:=SIZEOF(_handle),
					SRCADDR:=ADR(_handle),
					WRITE:=TRUE,
					TMOUT:=ADS_TIMEOUT);
				_state := 45;
			ELSE
				_state := 50;
			END_IF

		45: // wait for the release
			_releaseHandle(WRITE:=FALSE);
			IF NOT _releaseHandle.BUSY THEN
				THIS^.AssertFalse(_releaseHandle.ERR, 'Expected the symbol handle to be released');
				_hasHandle := FALSE;
				_state := 50;
			END_IF

		50: // done
			TcUnit.TEST_FINISHED();
	END_CASE
END_METHOD

END_FUNCTION_BLOCK

// ---- TEST/TRACING/SPAN/FB_TestSpan.TcPOU
(* Tests FB_Span.cloneTo, which processors use to keep a span that must outlive the original.
   A running span's context is taken through FB_Tracer.getSpanContext, tested in FB_TestTracer. *)
FUNCTION_BLOCK FB_TestSpan EXTENDS FB_TestSuite

THIS^.testCloneToCopiesEveryMember();
THIS^.testCloneToRejectsAssignedDestination();

(* cloneTo gives the copy its own copy of every member, so it outlives the source. *)
METHOD testCloneToCopiesEveryMember : REFERENCE TO FB_Test
VAR
	resource: FB_Resource('');
	idGenerator: FB_MockIdGenerator;
	provider: FB_TracerProvider_ForInspection(resource:=resource, idGenerator:=idGenerator, sampler:=TcOtlp_GVL.defaultSampler);
	scope: FB_InstrumentationScope('tracer.test', '1.0.0', '');
	tracer: FB_Tracer(scope:=scope, provider:=provider);
	pParent: POINTER TO FB_Span;
	pContext: POINTER TO FB_SpanContext;
	pSpan: POINTER TO FB_Span;
	pClone: POINTER TO FB_Span;
	pLink: POINTER TO FB_Link;
	pSourceLink: POINTER TO FB_Link;
	reason: E_SpanCloneFailureReason;
END_VAR
TcUnit.TEST('testCloneToCopiesEveryMember');
	IF resource.attributes.count = 0 THEN
		resource.attributes.setStringAttribute('host.id', 'PLC1');
	END_IF
	tracer.startSpan(name:='parent').build(pDest:=pParent);
	IF pParent <> 0 THEN tracer.getSpanContext(pSpan:=pParent, pDest:=pContext); END_IF
	tracer.startSpan(name:='work', kind:=E_SpanKind.SPAN_KIND_SERVER)
		.setParentUsingContext(pContext:=pContext)
		.addLink(pContext:=pContext)
		.setStringAttribute(key:='k', value:='v')
		.build(pDest:=pSpan);
	THIS^.AssertTrue(pSpan <> 0, 'Expected the span to build');
	IF pSpan <> 0 THEN
		// no builder sets timestamps; fixed values make the copy checkable
		pSpan^.startTimestamp := 1000;
		pSpan^.endTimestamp := 1500;
		tracer.setSpanStatusError(pSpan:=pSpan, message:='boom');
		pSpan^.links.reset();
		pSourceLink := pSpan^.links.next();

		THIS^.AssertTrue(pSpan^.cloneTo(pDest:=pClone, failureReason=>reason), 'Expected cloneTo to succeed');
		THIS^.AssertEquals_UDINT(TO_UDINT(E_SpanCloneFailureReason.NA), TO_UDINT(reason), 'Expected no failure');
		IF pClone <> 0 THEN
			THIS^.AssertTrue(pClone^.name <> 0 AND_THEN pClone^.name <> pSpan^.name, 'Expected a copied name');
			THIS^.AssertTrue(pClone^.traceId <> 0 AND_THEN pClone^.traceId <> pSpan^.traceId
				AND_THEN MEMCMP(ADR(pClone^.traceId^.bytes), ADR(pSpan^.traceId^.bytes), SIZEOF(pSpan^.traceId^.bytes)) = 0,
				'Expected a copied trace id');
			THIS^.AssertTrue(pClone^.spanId <> 0 AND_THEN pClone^.spanId <> pSpan^.spanId
				AND_THEN MEMCMP(ADR(pClone^.spanId^.bytes), ADR(pSpan^.spanId^.bytes), SIZEOF(pSpan^.spanId^.bytes)) = 0,
				'Expected a copied span id');
			THIS^.AssertTrue(pClone^.parentSpanId <> 0 AND_THEN pClone^.parentSpanId <> pSpan^.parentSpanId
				AND_THEN MEMCMP(ADR(pClone^.parentSpanId^.bytes), ADR(pSpan^.parentSpanId^.bytes), SIZEOF(pSpan^.parentSpanId^.bytes)) = 0,
				'Expected a copied parent span id');
			THIS^.AssertEquals_UDINT(TO_UDINT(E_SpanKind.SPAN_KIND_SERVER), TO_UDINT(pClone^.kind), 'Expected the kind');
			THIS^.AssertTrue(pClone^.startTimestamp = 1000 AND pClone^.endTimestamp = 1500, 'Expected the timestamps');
			THIS^.AssertEquals_UDINT(pSpan^.flags, pClone^.flags, 'Expected the flags');
			THIS^.AssertTrue(pClone^.status <> 0 AND_THEN pClone^.status <> pSpan^.status
				AND_THEN pClone^.status^.code = E_StatusCode.STATUS_CODE_ERROR
				AND_THEN pClone^.status^.message <> 0
				AND_THEN pClone^.status^.message <> pSpan^.status^.message,
				'Expected a copied error status');
			THIS^.AssertEquals_UDINT(pSpan^.attributes.count, pClone^.attributes.count, 'Expected the attributes');
			THIS^.AssertEquals_UDINT(1, pClone^.attributes.count, 'Expected one attribute');
			THIS^.AssertEquals_UDINT(1, pClone^.links.count, 'Expected one link');
			pClone^.links.reset();
			pLink := pClone^.links.next();
			THIS^.AssertTrue(pLink <> 0 AND_THEN pLink <> pSourceLink AND_THEN pLink^.spanId <> 0
				AND_THEN MEMCMP(ADR(pLink^.spanId^.bytes), ADR(pSourceLink^.spanId^.bytes), SIZEOF(pLink^.spanId^.bytes)) = 0,
				'Expected a copied link');
			THIS^.AssertEquals_UDINT(pSpan^.resource.attributes.count, pClone^.resource.attributes.count, 'Expected the resource');
			THIS^.AssertTrue(pClone^.resource.attributes.count > 0, 'Expected resource attributes to be copied');

			// the copy must stay valid once the source is gone
			pSpan^.delete(pSelf:=pSpan);
			THIS^.AssertEquals_STRING('work', pClone^.name^.pString^, 'Expected the name to outlive the source');
			THIS^.AssertEquals_STRING('boom', pClone^.status^.message^.pString^, 'Expected the message to outlive the source');
			pClone^.delete(pSelf:=pClone);
		END_IF
		IF pSpan <> 0 THEN pSpan^.delete(pSelf:=pSpan); END_IF
	END_IF
	IF pContext <> 0 THEN pContext^.delete(pSelf:=pContext); END_IF
	IF pParent <> 0 THEN pParent^.delete(pSelf:=pParent); END_IF
TcUnit.TEST_FINISHED();
END_METHOD

(* cloneTo refuses a destination that already holds a span and leaves it alone. *)
METHOD testCloneToRejectsAssignedDestination : REFERENCE TO FB_Test
VAR
	pSpan: POINTER TO FB_Span;
	pDest: POINTER TO FB_Span;
	reason: E_SpanCloneFailureReason;
END_VAR
TcUnit.TEST('testCloneToRejectsAssignedDestination');
	pSpan := __NEW(FB_Span);  // identity is irrelevant: only the destination check runs
	pDest := pSpan;  // deliberately assigned, so cloneTo must refuse it
	IF pSpan <> 0 THEN
		THIS^.AssertFalse(pSpan^.cloneTo(pDest:=pDest, failureReason=>reason), 'Expected cloneTo to fail');
		THIS^.AssertEquals_UDINT(
			TO_UDINT(E_SpanCloneFailureReason.DESTINATION_ALREADY_ASSIGNED),
			TO_UDINT(reason),
			'Expected DESTINATION_ALREADY_ASSIGNED'
		);
		THIS^.AssertTrue(pDest = pSpan, 'Expected the destination to be left alone');
		pSpan^.delete(pSelf:=pSpan);
	END_IF
TcUnit.TEST_FINISHED();
END_METHOD

END_FUNCTION_BLOCK

// ---- TEST/TRACING/PROVIDER/FB_TracerProvider_ForInspection.TcPOU
(* Provider test double that exposes the queue of ended spans for assertions. *)
FUNCTION_BLOCK FB_TracerProvider_ForInspection EXTENDS FB_TracerProvider

PROPERTY spans : REFERENCE TO FB_SpanQueue
GET
spans REF= THIS^._spans;
END_GET
END_PROPERTY

END_FUNCTION_BLOCK

// ---- TEST/TRACING/TRACER/FB_TestTracer.TcPOU
(* Tests the FB_Tracer fluent chain: validation at each step, identifier and flag assignment,
   and the hand-over of the built span to the caller. Also tests the methods that read and
   change a running span, which all refuse a null span. Each test builds its own provider and
   tracer around a deterministic id generator. *)
FUNCTION_BLOCK FB_TestTracer EXTENDS FB_TestSuite

THIS^.testBuildsRootSpan();
THIS^.testBuildsChildOfLocalParent();
THIS^.testChildOfRemoteParent();
THIS^.testRejectsInvalidParent();
THIS^.testBuildsChildOfSpan();
THIS^.testRejectsInvalidParentSpan();
THIS^.testKeepsFirstFailure();
THIS^.testRejectsEmptyName();
THIS^.testRejectsUnspecifiedKind();
THIS^.testBuildWithoutStartFails();
THIS^.testStartingSecondSpanFails();
THIS^.testBuildIntoAssignedDestinationFails();
THIS^.testNoIdentifiersAvailable();
THIS^.testSetsAttributes();
THIS^.testEndSpanQueuesSpan();
THIS^.testEndSpanRejectsNull();
THIS^.testEndSpanWithoutProcessorsQueuesSpan();
THIS^.testSetSpanStatusOk();
THIS^.testSetSpanStatusError();
THIS^.testSetSpanStatusFirstWins();
THIS^.testGetSpanContextCopiesIdentity();
THIS^.testGetSpanContextIsLocal();
THIS^.testGetSpanContextRejectsAssignedDestination();
THIS^.testGetSpanContextOnUnbuiltSpan();
THIS^.testAddsLinksToRunningSpan();
THIS^.testSetsRunningSpanAttributes();
THIS^.testDiscardSpanReleasesSpan();
THIS^.testRunningSpanMethodsRejectNullSpan();
THIS^.testAddsLinks();
THIS^.testRejectsInvalidLink();

(* A span without a parent starts a new trace: it gets fresh identifiers, no parent, root flags,
   and snapshots of the resource and scope. The tracer gives up ownership. *)
METHOD testBuildsRootSpan : REFERENCE TO FB_Test
VAR
	resource: FB_Resource('');
	idGenerator: FB_MockIdGenerator;
	provider: FB_TracerProvider(resource:=resource, idGenerator:=idGenerator, sampler:=TcOtlp_GVL.defaultSampler);
	scope: FB_InstrumentationScope('tracer.test', '1.0.0', '');
	tracer: FB_Tracer(scope:=scope, provider:=provider);
	pSpan: POINTER TO FB_Span;
	success: BOOL;
	reason: E_TracerFailureReason;
END_VAR
TcUnit.TEST('testBuildsRootSpan');
	success := tracer.startSpan(name:='root').build(pDest:=pSpan, failureReason=>reason);
	THIS^.AssertTrue(success, 'Expected a root span to build');
	THIS^.AssertEquals_UDINT(
		TO_UDINT(E_TracerFailureReason.NA),
		TO_UDINT(reason),
		'Expected no failure reason on success'
	);
	THIS^.AssertTrue(pSpan <> 0, 'Expected build to assign the destination');
	THIS^.AssertTrue(tracer.pSpan = 0, 'Expected the tracer to hand over the span');

	IF pSpan <> 0 THEN
		THIS^.AssertTrue(pSpan^.traceId <> 0, 'Expected a trace id');
		THIS^.AssertTrue(pSpan^.spanId <> 0, 'Expected a span id');
		THIS^.AssertTrue(pSpan^.parentSpanId = 0, 'Expected a root span to have no parent');
		THIS^.AssertTrue(pSpan^.traceState = 0, 'Expected a root span to have no trace state');
		THIS^.AssertTrue(pSpan^.name <> 0, 'Expected a name');
		IF pSpan^.name <> 0 THEN
			THIS^.AssertEquals_STRING('root', pSpan^.name^.pString^, 'Expected the name to be copied');
		END_IF
		THIS^.AssertEquals_UDINT(
			TO_UDINT(E_SpanKind.SPAN_KIND_INTERNAL),
			TO_UDINT(pSpan^.kind),
			'Expected the default kind to be INTERNAL'
		);
		THIS^.AssertTrue(pSpan^.startTimestamp > 0, 'Expected a start timestamp');
		THIS^.AssertEquals_UDINT(16#101, pSpan^.flags, 'Expected a root span to be sampled with remoteness known');
		THIS^.AssertEquals_STRING('tracer.test', pSpan^.scope.name, 'Expected the scope to be snapshotted');
		pSpan^.delete(pSelf:=pSpan);
	END_IF
TcUnit.TEST_FINISHED();
END_METHOD

(* A child of a local span continues its trace, records the parent's span id, and takes its
   own span id. *)
METHOD testBuildsChildOfLocalParent : REFERENCE TO FB_Test
VAR
	resource: FB_Resource('');
	idGenerator: FB_MockIdGenerator;
	provider: FB_TracerProvider(resource:=resource, idGenerator:=idGenerator, sampler:=TcOtlp_GVL.defaultSampler);
	scope: FB_InstrumentationScope('tracer.test', '1.0.0', '');
	tracer: FB_Tracer(scope:=scope, provider:=provider);
	pRoot: POINTER TO FB_Span;
	pChild: POINTER TO FB_Span;
	pContext: POINTER TO FB_SpanContext;
	success: BOOL;
	reason: E_TracerFailureReason;
END_VAR
TcUnit.TEST('testBuildsChildOfLocalParent');
	tracer.startSpan(name:='root').build(pDest:=pRoot);
	IF pRoot <> 0 THEN
		tracer.getSpanContext(pSpan:=pRoot, pDest:=pContext);
	END_IF

	success := tracer
		.startSpan(name:='child', kind:=E_SpanKind.SPAN_KIND_CLIENT)
		.setParentUsingContext(pContext:=pContext)
		.build(pDest:=pChild, failureReason=>reason);
	THIS^.AssertTrue(success, 'Expected a child span to build');
	THIS^.AssertEquals_UDINT(
		TO_UDINT(E_TracerFailureReason.NA),
		TO_UDINT(reason),
		'Expected no failure reason on success'
	);

	IF pRoot <> 0 AND_THEN pChild <> 0 THEN
		THIS^.AssertTrue(
			MEMCMP(ADR(pChild^.traceId^.bytes), ADR(pRoot^.traceId^.bytes), SIZEOF(pRoot^.traceId^.bytes)) = 0,
			'Expected the child to continue the parent$'s trace'
		);
		THIS^.AssertTrue(pChild^.parentSpanId <> 0, 'Expected the child to record its parent');
		IF pChild^.parentSpanId <> 0 THEN
			THIS^.AssertTrue(
				MEMCMP(ADR(pChild^.parentSpanId^.bytes), ADR(pRoot^.spanId^.bytes), SIZEOF(pRoot^.spanId^.bytes)) = 0,
				'Expected the parent span id to be the root$'s span id'
			);
		END_IF
		THIS^.AssertTrue(
			MEMCMP(ADR(pChild^.spanId^.bytes), ADR(pRoot^.spanId^.bytes), SIZEOF(pRoot^.spanId^.bytes)) <> 0,
			'Expected the child to have its own span id'
		);
		THIS^.AssertEquals_UDINT(16#101, pChild^.flags, 'Expected a local parent to set bit 8 but not bit 9');
		THIS^.AssertEquals_UDINT(
			TO_UDINT(E_SpanKind.SPAN_KIND_CLIENT),
			TO_UDINT(pChild^.kind),
			'Expected the kind to be kept'
		);
	END_IF

	IF pContext <> 0 THEN pContext^.delete(pSelf:=pContext); END_IF
	IF pChild <> 0 THEN pChild^.delete(pSelf:=pChild); END_IF
	IF pRoot <> 0 THEN pRoot^.delete(pSelf:=pRoot); END_IF
TcUnit.TEST_FINISHED();
END_METHOD

(* A remote parent sets bits 8 and 9 on the child and its trace state is copied. The child's
   own context is still local. *)
METHOD testChildOfRemoteParent : REFERENCE TO FB_Test
VAR
	resource: FB_Resource('');
	idGenerator: FB_MockIdGenerator;
	provider: FB_TracerProvider(resource:=resource, idGenerator:=idGenerator, sampler:=TcOtlp_GVL.defaultSampler);
	scope: FB_InstrumentationScope('tracer.test', '1.0.0', '');
	tracer: FB_Tracer(scope:=scope, provider:=provider);
	pChild: POINTER TO FB_Span;
	pRemote: POINTER TO FB_SpanContext;
	pChildContext: POINTER TO FB_SpanContext;
	traceId: FB_TraceId;
	spanId: FB_SpanId;
	traceStateText: T_MaxString := 'vendor=abc';
	pTraceState: POINTER TO FB_TraceState;
	success: BOOL;
	reason: E_TracerFailureReason;
END_VAR
TcUnit.TEST('testChildOfRemoteParent');
	MEMSET(ADR(traceId.bytes), 16#AA, SIZEOF(traceId.bytes));
	MEMSET(ADR(spanId.bytes), 16#BB, SIZEOF(spanId.bytes));
	TraceStateFactory.parse(pDest:=pTraceState, pHeader:=ADR(traceStateText));
	ContextFactory.buildContext(
		pDest:=pRemote,
		pTraceId:=ADR(traceId),
		pSpanId:=ADR(spanId),
		pTraceState:=pTraceState,
		traceFlags:=16#301
	);
	IF pTraceState <> 0 THEN pTraceState^.delete(pSelf:=pTraceState); END_IF

	success := tracer
		.startSpan(name:='remote.child', kind:=E_SpanKind.SPAN_KIND_CONSUMER)
		.setParentUsingContext(pContext:=pRemote)
		.build(pDest:=pChild, failureReason=>reason);
	THIS^.AssertTrue(success, 'Expected a child of a remote parent to build');
	THIS^.AssertEquals_UDINT(
		TO_UDINT(E_TracerFailureReason.NA),
		TO_UDINT(reason),
		'Expected no failure reason on success'
	);

	// the context is borrowed, so it can be released before the span
	IF pRemote <> 0 THEN pRemote^.delete(pSelf:=pRemote); END_IF

	IF pChild <> 0 THEN
		THIS^.AssertEquals_UDINT(16#301, pChild^.flags, 'Expected a remote parent to set bits 8 and 9');
		THIS^.AssertTrue(
			MEMCMP(ADR(pChild^.traceId^.bytes), ADR(traceId.bytes), SIZEOF(traceId.bytes)) = 0,
			'Expected the child to continue the remote trace'
		);
		THIS^.AssertTrue(pChild^.traceState <> 0, 'Expected the trace state to be copied');
		IF pChild^.traceState <> 0 THEN
			THIS^.AssertEquals_STRING('vendor=abc', pChild^.traceState^.pString^, 'Expected the trace state text to be copied');
		END_IF

		tracer.getSpanContext(pSpan:=pChild, pDest:=pChildContext);
		THIS^.AssertTrue(pChildContext <> 0, 'Expected a context from the child');
		IF pChildContext <> 0 THEN
			THIS^.AssertFalse(pChildContext^.isRemote(), 'Expected the child$'s own context to be local');
			THIS^.AssertEquals_UDINT(16#101, pChildContext^.traceFlags, 'Expected the sampled bit and bit 8 only');
			pChildContext^.delete(pSelf:=pChildContext);
		END_IF
		pChild^.delete(pSelf:=pChild);
	END_IF
TcUnit.TEST_FINISHED();
END_METHOD

(* A parent context with all zero identifiers is rejected and nothing is handed over. *)
METHOD testRejectsInvalidParent : REFERENCE TO FB_Test
VAR
	resource: FB_Resource('');
	idGenerator: FB_MockIdGenerator;
	provider: FB_TracerProvider(resource:=resource, idGenerator:=idGenerator, sampler:=TcOtlp_GVL.defaultSampler);
	scope: FB_InstrumentationScope('tracer.test', '1.0.0', '');
	tracer: FB_Tracer(scope:=scope, provider:=provider);
	pSpan: POINTER TO FB_Span;
	pContext: POINTER TO FB_SpanContext;
	traceId: FB_TraceId;
	spanId: FB_SpanId;
	success: BOOL;
	reason: E_TracerFailureReason;
END_VAR
TcUnit.TEST('testRejectsInvalidParent');
	ContextFactory.buildContext(pDest:=pContext, pTraceId:=ADR(traceId), pSpanId:=ADR(spanId), pTraceState:=0, traceFlags:=16#101);

	success := tracer.startSpan(name:='child').setParentUsingContext(pContext:=pContext).build(pDest:=pSpan, failureReason=>reason);
	THIS^.AssertFalse(success, 'Expected an invalid parent to fail the chain');
	THIS^.AssertEquals_UDINT(
		TO_UDINT(E_TracerFailureReason.PARENT_CONTEXT_INVALID),
		TO_UDINT(reason),
		'Expected PARENT_CONTEXT_INVALID'
	);
	THIS^.AssertTrue(pSpan = 0, 'Expected the destination to stay unassigned');
	THIS^.AssertTrue(tracer.pSpan = 0, 'Expected the incomplete span to be released');

	IF pContext <> 0 THEN pContext^.delete(pSelf:=pContext); END_IF
	IF pSpan <> 0 THEN pSpan^.delete(pSelf:=pSpan); END_IF
TcUnit.TEST_FINISHED();
END_METHOD

(* setParentUsingSpan takes the parent's identity straight from a built span: the child
   continues its trace, records its span id, copies its trace state and marks the parent as
   local, even when the parent itself has a remote parent. *)
METHOD testBuildsChildOfSpan : REFERENCE TO FB_Test
VAR
	resource: FB_Resource('');
	idGenerator: FB_MockIdGenerator;
	provider: FB_TracerProvider(resource:=resource, idGenerator:=idGenerator, sampler:=TcOtlp_GVL.defaultSampler);
	scope: FB_InstrumentationScope('tracer.test', '1.0.0', '');
	tracer: FB_Tracer(scope:=scope, provider:=provider);
	pRemote: POINTER TO FB_SpanContext;
	pParent: POINTER TO FB_Span;
	pChild: POINTER TO FB_Span;
	traceId: FB_TraceId;
	spanId: FB_SpanId;
	traceStateText: T_MaxString := 'vendor=abc';
	pTraceState: POINTER TO FB_TraceState;
	success: BOOL;
	reason: E_TracerFailureReason;
END_VAR
TcUnit.TEST('testBuildsChildOfSpan');
	MEMSET(ADR(traceId.bytes), 16#AA, SIZEOF(traceId.bytes));
	MEMSET(ADR(spanId.bytes), 16#BB, SIZEOF(spanId.bytes));
	TraceStateFactory.parse(pDest:=pTraceState, pHeader:=ADR(traceStateText));
	ContextFactory.buildContext(
		pDest:=pRemote,
		pTraceId:=ADR(traceId),
		pSpanId:=ADR(spanId),
		pTraceState:=pTraceState,
		traceFlags:=16#301
	);
	IF pTraceState <> 0 THEN pTraceState^.delete(pSelf:=pTraceState); END_IF
	tracer.startSpan(name:='parent').setParentUsingContext(pContext:=pRemote).build(pDest:=pParent);
	IF pRemote <> 0 THEN pRemote^.delete(pSelf:=pRemote); END_IF
	THIS^.AssertTrue(pParent <> 0, 'Expected the parent span to build');

	success := tracer
		.startSpan(name:='child')
		.setParentUsingSpan(pParentSpan:=pParent)
		.build(pDest:=pChild, failureReason=>reason);
	THIS^.AssertTrue(success, 'Expected a child of a span to build');
	THIS^.AssertEquals_UDINT(
		TO_UDINT(E_TracerFailureReason.NA),
		TO_UDINT(reason),
		'Expected no failure reason on success'
	);

	IF pParent <> 0 AND_THEN pChild <> 0 THEN
		THIS^.AssertTrue(
			MEMCMP(ADR(pChild^.traceId^.bytes), ADR(pParent^.traceId^.bytes), SIZEOF(pParent^.traceId^.bytes)) = 0,
			'Expected the child to continue the parent$'s trace'
		);
		THIS^.AssertTrue(pChild^.parentSpanId <> 0, 'Expected the child to record its parent');
		IF pChild^.parentSpanId <> 0 THEN
			THIS^.AssertTrue(
				MEMCMP(ADR(pChild^.parentSpanId^.bytes), ADR(pParent^.spanId^.bytes), SIZEOF(pParent^.spanId^.bytes)) = 0,
				'Expected the parent span id to be the parent$'s span id'
			);
		END_IF
		THIS^.AssertEquals_UDINT(16#101, pChild^.flags, 'Expected a span parent to be local: bit 8 set, bit 9 clear');
		THIS^.AssertTrue(pChild^.traceState <> 0, 'Expected the trace state to be copied');
		IF pChild^.traceState <> 0 THEN
			THIS^.AssertTrue(pChild^.traceState <> pParent^.traceState, 'Expected the child to own its own trace state');
			THIS^.AssertEquals_STRING('vendor=abc', pChild^.traceState^.pString^, 'Expected the trace state text to be copied');
		END_IF
	END_IF

	IF pChild <> 0 THEN pChild^.delete(pSelf:=pChild); END_IF
	IF pParent <> 0 THEN pParent^.delete(pSelf:=pParent); END_IF
TcUnit.TEST_FINISHED();
END_METHOD

(* setParentUsingSpan refuses a null span and a span that has not been built, and nothing is
   handed over. *)
METHOD testRejectsInvalidParentSpan : REFERENCE TO FB_Test
VAR
	resource: FB_Resource('');
	idGenerator: FB_MockIdGenerator;
	provider: FB_TracerProvider(resource:=resource, idGenerator:=idGenerator, sampler:=TcOtlp_GVL.defaultSampler);
	scope: FB_InstrumentationScope('tracer.test', '1.0.0', '');
	tracer: FB_Tracer(scope:=scope, provider:=provider);
	unbuilt: FB_Span;
	pSpan: POINTER TO FB_Span;
	success: BOOL;
	reason: E_TracerFailureReason;
END_VAR
TcUnit.TEST('testRejectsInvalidParentSpan');
	success := tracer.startSpan(name:='child').setParentUsingSpan(pParentSpan:=0).build(pDest:=pSpan, failureReason=>reason);
	THIS^.AssertFalse(success, 'Expected a null parent span to fail the chain');
	THIS^.AssertEquals_UDINT(
		TO_UDINT(E_TracerFailureReason.PARENT_SPAN_POINTER_NULL),
		TO_UDINT(reason),
		'Expected PARENT_SPAN_POINTER_NULL'
	);
	THIS^.AssertTrue(pSpan = 0, 'Expected the destination to stay unassigned');

	success := tracer.startSpan(name:='child').setParentUsingSpan(pParentSpan:=ADR(unbuilt)).build(pDest:=pSpan, failureReason=>reason);
	THIS^.AssertFalse(success, 'Expected a parent span without identifiers to fail the chain');
	THIS^.AssertEquals_UDINT(
		TO_UDINT(E_TracerFailureReason.PARENT_SPAN_INVALID),
		TO_UDINT(reason),
		'Expected PARENT_SPAN_INVALID'
	);
	THIS^.AssertTrue(pSpan = 0, 'Expected the destination to stay unassigned');
	THIS^.AssertTrue(tracer.pSpan = 0, 'Expected the incomplete span to be released');

	IF pSpan <> 0 THEN pSpan^.delete(pSelf:=pSpan); END_IF
TcUnit.TEST_FINISHED();
END_METHOD

(* Later steps in a failed chain do not replace the first failure. *)
METHOD testKeepsFirstFailure : REFERENCE TO FB_Test
VAR
	resource: FB_Resource('');
	idGenerator: FB_MockIdGenerator;
	provider: FB_TracerProvider(resource:=resource, idGenerator:=idGenerator, sampler:=TcOtlp_GVL.defaultSampler);
	scope: FB_InstrumentationScope('tracer.test', '1.0.0', '');
	tracer: FB_Tracer(scope:=scope, provider:=provider);
	pSpan: POINTER TO FB_Span;
	success: BOOL;
	reason: E_TracerFailureReason;
END_VAR
TcUnit.TEST('testKeepsFirstFailure');
	success := tracer
		.startSpan(name:='child')
		.setParentUsingContext(pContext:=0)
		.setStringAttribute('key', 'value')
		.build(pDest:=pSpan, failureReason=>reason);
	THIS^.AssertFalse(success, 'Expected a null parent to fail the chain');
	THIS^.AssertEquals_UDINT(
		TO_UDINT(E_TracerFailureReason.PARENT_CONTEXT_POINTER_NULL),
		TO_UDINT(reason),
		'Expected the first failure to be reported'
	);
	THIS^.AssertTrue(pSpan = 0, 'Expected the destination to stay unassigned');

	// the failure does not carry over to the next chain
	success := tracer.startSpan(name:='next').build(pDest:=pSpan, failureReason=>reason);
	THIS^.AssertTrue(success, 'Expected the next chain to start clean');
	IF pSpan <> 0 THEN pSpan^.delete(pSelf:=pSpan); END_IF
TcUnit.TEST_FINISHED();
END_METHOD

(* OTLP requires a span name. *)
METHOD testRejectsEmptyName : REFERENCE TO FB_Test
VAR
	resource: FB_Resource('');
	idGenerator: FB_MockIdGenerator;
	provider: FB_TracerProvider(resource:=resource, idGenerator:=idGenerator, sampler:=TcOtlp_GVL.defaultSampler);
	scope: FB_InstrumentationScope('tracer.test', '1.0.0', '');
	tracer: FB_Tracer(scope:=scope, provider:=provider);
	pSpan: POINTER TO FB_Span;
	success: BOOL;
	reason: E_TracerFailureReason;
END_VAR
TcUnit.TEST('testRejectsEmptyName');
	success := tracer.startSpan(name:='').build(pDest:=pSpan, failureReason=>reason);
	THIS^.AssertFalse(success, 'Expected an empty name to fail');
	THIS^.AssertEquals_UDINT(
		TO_UDINT(E_TracerFailureReason.SPAN_NAME_EMPTY),
		TO_UDINT(reason),
		'Expected SPAN_NAME_EMPTY'
	);
	THIS^.AssertTrue(pSpan = 0, 'Expected the destination to stay unassigned');
	IF pSpan <> 0 THEN pSpan^.delete(pSelf:=pSpan); END_IF
TcUnit.TEST_FINISHED();
END_METHOD

(* OTLP says SPAN_KIND_UNSPECIFIED must not be used. *)
METHOD testRejectsUnspecifiedKind : REFERENCE TO FB_Test
VAR
	resource: FB_Resource('');
	idGenerator: FB_MockIdGenerator;
	provider: FB_TracerProvider(resource:=resource, idGenerator:=idGenerator, sampler:=TcOtlp_GVL.defaultSampler);
	scope: FB_InstrumentationScope('tracer.test', '1.0.0', '');
	tracer: FB_Tracer(scope:=scope, provider:=provider);
	pSpan: POINTER TO FB_Span;
	success: BOOL;
	reason: E_TracerFailureReason;
END_VAR
TcUnit.TEST('testRejectsUnspecifiedKind');
	success := tracer.startSpan(name:='span', kind:=E_SpanKind.SPAN_KIND_UNSPECIFIED).build(pDest:=pSpan, failureReason=>reason);
	THIS^.AssertFalse(success, 'Expected an unspecified kind to fail');
	THIS^.AssertEquals_UDINT(
		TO_UDINT(E_TracerFailureReason.SPAN_KIND_UNSPECIFIED),
		TO_UDINT(reason),
		'Expected SPAN_KIND_UNSPECIFIED'
	);
	THIS^.AssertTrue(pSpan = 0, 'Expected the destination to stay unassigned');
	IF pSpan <> 0 THEN pSpan^.delete(pSelf:=pSpan); END_IF
TcUnit.TEST_FINISHED();
END_METHOD

(* build and the setters need a span that startSpan created. *)
METHOD testBuildWithoutStartFails : REFERENCE TO FB_Test
VAR
	resource: FB_Resource('');
	idGenerator: FB_MockIdGenerator;
	provider: FB_TracerProvider(resource:=resource, idGenerator:=idGenerator, sampler:=TcOtlp_GVL.defaultSampler);
	scope: FB_InstrumentationScope('tracer.test', '1.0.0', '');
	tracer: FB_Tracer(scope:=scope, provider:=provider);
	pSpan: POINTER TO FB_Span;
	success: BOOL;
	reason: E_TracerFailureReason;
END_VAR
TcUnit.TEST('testBuildWithoutStartFails');
	success := tracer.setStringAttribute('key', 'value').build(pDest:=pSpan, failureReason=>reason);
	THIS^.AssertFalse(success, 'Expected build without startSpan to fail');
	THIS^.AssertEquals_UDINT(
		TO_UDINT(E_TracerFailureReason.SPAN_NOT_STARTED),
		TO_UDINT(reason),
		'Expected SPAN_NOT_STARTED'
	);
	THIS^.AssertTrue(pSpan = 0, 'Expected the destination to stay unassigned');
TcUnit.TEST_FINISHED();
END_METHOD

(* The tracer builds one span at a time. A second startSpan fails the chain, and build
   releases the span that was already building. *)
METHOD testStartingSecondSpanFails : REFERENCE TO FB_Test
VAR
	resource: FB_Resource('');
	idGenerator: FB_MockIdGenerator;
	provider: FB_TracerProvider(resource:=resource, idGenerator:=idGenerator, sampler:=TcOtlp_GVL.defaultSampler);
	scope: FB_InstrumentationScope('tracer.test', '1.0.0', '');
	tracer: FB_Tracer(scope:=scope, provider:=provider);
	pSpan: POINTER TO FB_Span;
	success: BOOL;
	reason: E_TracerFailureReason;
END_VAR
TcUnit.TEST('testStartingSecondSpanFails');
	tracer.startSpan(name:='first');
	success := tracer.startSpan(name:='second').build(pDest:=pSpan, failureReason=>reason);
	THIS^.AssertFalse(success, 'Expected a second startSpan to fail');
	THIS^.AssertEquals_UDINT(
		TO_UDINT(E_TracerFailureReason.SPAN_ALREADY_STARTED),
		TO_UDINT(reason),
		'Expected SPAN_ALREADY_STARTED'
	);
	THIS^.AssertTrue(pSpan = 0, 'Expected the destination to stay unassigned');
	THIS^.AssertTrue(tracer.pSpan = 0, 'Expected build to release the building span');
	IF pSpan <> 0 THEN pSpan^.delete(pSelf:=pSpan); END_IF
TcUnit.TEST_FINISHED();
END_METHOD

(* build follows the VAR_IN_OUT pointer pattern: it never overwrites a span the caller owns. *)
METHOD testBuildIntoAssignedDestinationFails : REFERENCE TO FB_Test
VAR
	resource: FB_Resource('');
	idGenerator: FB_MockIdGenerator;
	provider: FB_TracerProvider(resource:=resource, idGenerator:=idGenerator, sampler:=TcOtlp_GVL.defaultSampler);
	scope: FB_InstrumentationScope('tracer.test', '1.0.0', '');
	tracer: FB_Tracer(scope:=scope, provider:=provider);
	pSpan: POINTER TO FB_Span;
	pFirst: POINTER TO FB_Span;
	success: BOOL;
	reason: E_TracerFailureReason;
END_VAR
TcUnit.TEST('testBuildIntoAssignedDestinationFails');
	tracer.startSpan(name:='first').build(pDest:=pSpan);
	pFirst := pSpan;

	success := tracer.startSpan(name:='second').build(pDest:=pSpan, failureReason=>reason);
	THIS^.AssertFalse(success, 'Expected build into an assigned destination to fail');
	THIS^.AssertEquals_UDINT(
		TO_UDINT(E_TracerFailureReason.DESTINATION_ALREADY_ASSIGNED),
		TO_UDINT(reason),
		'Expected DESTINATION_ALREADY_ASSIGNED'
	);
	THIS^.AssertTrue(pSpan = pFirst, 'Expected the destination pointer to be left alone');
	THIS^.AssertTrue(tracer.pSpan = 0, 'Expected the second span to be released');
	IF pSpan <> 0 THEN pSpan^.delete(pSelf:=pSpan); END_IF
TcUnit.TEST_FINISHED();
END_METHOD

(* A generator with nothing ready fails the build with a retryable reason. *)
METHOD testNoIdentifiersAvailable : REFERENCE TO FB_Test
VAR
	resource: FB_Resource('');
	idGenerator: FB_MockIdGenerator;
	provider: FB_TracerProvider(resource:=resource, idGenerator:=idGenerator, sampler:=TcOtlp_GVL.defaultSampler);
	scope: FB_InstrumentationScope('tracer.test', '1.0.0', '');
	tracer: FB_Tracer(scope:=scope, provider:=provider);
	pSpan: POINTER TO FB_Span;
	success: BOOL;
	reason: E_TracerFailureReason;
END_VAR
TcUnit.TEST('testNoIdentifiersAvailable');
	idGenerator.available := FALSE;
	success := tracer.startSpan(name:='root').build(pDest:=pSpan, failureReason=>reason);
	THIS^.AssertFalse(success, 'Expected build to fail without identifiers');
	THIS^.AssertEquals_UDINT(
		TO_UDINT(E_TracerFailureReason.IDENTIFIERS_UNAVAILABLE),
		TO_UDINT(reason),
		'Expected IDENTIFIERS_UNAVAILABLE'
	);
	THIS^.AssertTrue(pSpan = 0, 'Expected the destination to stay unassigned');
	THIS^.AssertTrue(tracer.pSpan = 0, 'Expected the incomplete span to be released');
	IF pSpan <> 0 THEN pSpan^.delete(pSelf:=pSpan); END_IF
TcUnit.TEST_FINISHED();
END_METHOD

(* Attributes set during the chain are owned by the built span. *)
METHOD testSetsAttributes : REFERENCE TO FB_Test
VAR
	resource: FB_Resource('');
	idGenerator: FB_MockIdGenerator;
	provider: FB_TracerProvider(resource:=resource, idGenerator:=idGenerator, sampler:=TcOtlp_GVL.defaultSampler);
	scope: FB_InstrumentationScope('tracer.test', '1.0.0', '');
	tracer: FB_Tracer(scope:=scope, provider:=provider);
	pSpan: POINTER TO FB_Span;
	setpoint: DINT := 42;
	success: BOOL;
	reason: E_TracerFailureReason;
END_VAR
TcUnit.TEST('testSetsAttributes');
	success := tracer
		.startSpan(name:='span')
		.setStringAttribute('skid', 'A')
		.setNumberAttribute('setpoint', setpoint)
		.build(pDest:=pSpan, failureReason=>reason);
	THIS^.AssertTrue(success, 'Expected a span with attributes to build');
	THIS^.AssertEquals_UDINT(
		TO_UDINT(E_TracerFailureReason.NA),
		TO_UDINT(reason),
		'Expected no failure reason on success'
	);
	IF pSpan <> 0 THEN
		THIS^.AssertEquals_UDINT(2, pSpan^.attributes.count, 'Expected both attributes on the span');
		pSpan^.delete(pSelf:=pSpan);
	END_IF
TcUnit.TEST_FINISHED();
END_METHOD

(* endSpan stamps the end time, moves the span into the provider's queue, and clears the
   caller's pointer. *)
METHOD testEndSpanQueuesSpan : REFERENCE TO FB_Test
VAR
	resource: FB_Resource('');
	idGenerator: FB_MockIdGenerator;
	provider: FB_TracerProvider_ForInspection(resource:=resource, idGenerator:=idGenerator, sampler:=TcOtlp_GVL.defaultSampler);
	scope: FB_InstrumentationScope('tracer.test', '1.0.0', '');
	tracer: FB_Tracer(scope:=scope, provider:=provider);
	processor: FB_SpanProcessor_ForInspection(exporter:=0);
	pSpan: POINTER TO FB_Span;
	pExpected: POINTER TO FB_Span;
	pEnded: POINTER TO FB_Span;
	success: BOOL;
	reason: E_TracerFailureReason;
	queueReason: E_SpanQueueFailureReason;
END_VAR
TcUnit.TEST('testEndSpanQueuesSpan');
	provider.stageProcessor(processor);
	success := tracer.startSpan(name:='work').build(pDest:=pSpan, failureReason=>reason);
	THIS^.AssertTrue(success, 'Expected the span to build');
	pExpected := pSpan;

	success := tracer.endSpan(pSpan:=pSpan, failureReason=>reason);
	THIS^.AssertTrue(success, 'Expected endSpan to succeed');
	THIS^.AssertEquals_UDINT(
		TO_UDINT(E_TracerFailureReason.NA),
		TO_UDINT(reason),
		'Expected no failure reason on success'
	);
	THIS^.AssertTrue(pSpan = 0, 'Expected endSpan to clear the caller$'s pointer');
	THIS^.AssertEquals_UDINT(1, provider.spans.count, 'Expected the provider to queue the span');

	provider.spans.pop(pValue:=pEnded, failureReason=>queueReason);
	THIS^.AssertTrue(pEnded = pExpected, 'Expected the queued span to be the one that was ended');
	IF pEnded <> 0 THEN
		THIS^.AssertTrue(pEnded^.endTimestamp <> 0, 'Expected an end timestamp');
		THIS^.AssertTrue(
			pEnded^.endTimestamp >= pEnded^.startTimestamp,
			'Expected the span to end no earlier than it started'
		);
		pEnded^.delete(pSelf:=pEnded);
	END_IF
	IF pSpan <> 0 THEN pSpan^.delete(pSelf:=pSpan); END_IF
TcUnit.TEST_FINISHED();
END_METHOD

(* A null span pointer is refused and nothing is queued. *)
METHOD testEndSpanRejectsNull : REFERENCE TO FB_Test
VAR
	resource: FB_Resource('');
	idGenerator: FB_MockIdGenerator;
	provider: FB_TracerProvider_ForInspection(resource:=resource, idGenerator:=idGenerator, sampler:=TcOtlp_GVL.defaultSampler);
	scope: FB_InstrumentationScope('tracer.test', '1.0.0', '');
	tracer: FB_Tracer(scope:=scope, provider:=provider);
	pSpan: POINTER TO FB_Span;
	success: BOOL;
	reason: E_TracerFailureReason;
END_VAR
TcUnit.TEST('testEndSpanRejectsNull');
	success := tracer.endSpan(pSpan:=pSpan, failureReason=>reason);
	THIS^.AssertFalse(success, 'Expected endSpan to fail without a span');
	THIS^.AssertEquals_UDINT(
		TO_UDINT(E_TracerFailureReason.SPAN_POINTER_NULL),
		TO_UDINT(reason),
		'Expected SPAN_POINTER_NULL'
	);
	THIS^.AssertEquals_UDINT(0, provider.spans.count, 'Expected nothing to be queued');
TcUnit.TEST_FINISHED();
END_METHOD

(* With no processor staged yet, endSpan still queues the span for the provider's next tick. *)
METHOD testEndSpanWithoutProcessorsQueuesSpan : REFERENCE TO FB_Test
VAR
	resource: FB_Resource('');
	idGenerator: FB_MockIdGenerator;
	provider: FB_TracerProvider_ForInspection(resource:=resource, idGenerator:=idGenerator, sampler:=TcOtlp_GVL.defaultSampler);
	scope: FB_InstrumentationScope('tracer.test', '1.0.0', '');
	tracer: FB_Tracer(scope:=scope, provider:=provider);
	pSpan: POINTER TO FB_Span;
	success: BOOL;
	reason: E_TracerFailureReason;
END_VAR
TcUnit.TEST('testEndSpanWithoutProcessorsQueuesSpan');
	tracer.startSpan(name:='work').build(pDest:=pSpan);
	THIS^.AssertTrue(pSpan <> 0, 'Expected the span to build');

	success := tracer.endSpan(pSpan:=pSpan, failureReason=>reason);
	THIS^.AssertTrue(success, 'Expected endSpan to succeed');
	THIS^.AssertEquals_UDINT(
		TO_UDINT(E_TracerFailureReason.NA),
		TO_UDINT(reason),
		'Expected no failure reason'
	);
	THIS^.AssertTrue(pSpan = 0, 'Expected endSpan to clear the caller$'s pointer');
	THIS^.AssertEquals_UDINT(1, provider.spans.count, 'Expected the span to be queued');
	IF pSpan <> 0 THEN pSpan^.delete(pSelf:=pSpan); END_IF
TcUnit.TEST_FINISHED();
END_METHOD

(* setSpanStatusOk gives a span with no status an OK status without a message. *)
METHOD testSetSpanStatusOk : REFERENCE TO FB_Test
VAR
	resource: FB_Resource('');
	idGenerator: FB_MockIdGenerator;
	provider: FB_TracerProvider(resource:=resource, idGenerator:=idGenerator, sampler:=TcOtlp_GVL.defaultSampler);
	scope: FB_InstrumentationScope('tracer.test', '1.0.0', '');
	tracer: FB_Tracer(scope:=scope, provider:=provider);
	span: FB_Span;  // a bare span: the status setters need no identity
	success: BOOL;
	reason: E_TracerFailureReason;
END_VAR
TcUnit.TEST('testSetSpanStatusOk');
	success := tracer.setSpanStatusOk(pSpan:=ADR(span), failureReason=>reason);
	THIS^.AssertTrue(success, 'Expected setSpanStatusOk to succeed');
	THIS^.AssertEquals_UDINT(TO_UDINT(E_TracerFailureReason.NA), TO_UDINT(reason), 'Expected no failure');
	THIS^.AssertTrue(span.status <> 0, 'Expected a status');
	IF span.status <> 0 THEN
		THIS^.AssertEquals_UDINT(TO_UDINT(E_StatusCode.STATUS_CODE_OK), TO_UDINT(span.status^.code), 'Expected an OK code');
		THIS^.AssertTrue(span.status^.message = 0, 'Expected no message');
	END_IF
	span.free();
TcUnit.TEST_FINISHED();
END_METHOD

(* setSpanStatusError keeps its own copy of the message, and an empty message leaves the
   status without one. *)
METHOD testSetSpanStatusError : REFERENCE TO FB_Test
VAR
	resource: FB_Resource('');
	idGenerator: FB_MockIdGenerator;
	provider: FB_TracerProvider(resource:=resource, idGenerator:=idGenerator, sampler:=TcOtlp_GVL.defaultSampler);
	scope: FB_InstrumentationScope('tracer.test', '1.0.0', '');
	tracer: FB_Tracer(scope:=scope, provider:=provider);
	span: FB_Span;  // a bare span: the status setters need no identity
	emptySpan: FB_Span;
	message: T_MaxString := 'motor over temp';
	success: BOOL;
	reason: E_TracerFailureReason;
END_VAR
TcUnit.TEST('testSetSpanStatusError');
	success := tracer.setSpanStatusError(pSpan:=ADR(span), message:=message, failureReason=>reason);
	message := 'changed by the caller';
	THIS^.AssertTrue(success, 'Expected setSpanStatusError to succeed');
	THIS^.AssertEquals_UDINT(TO_UDINT(E_TracerFailureReason.NA), TO_UDINT(reason), 'Expected no failure');
	THIS^.AssertTrue(span.status <> 0, 'Expected a status');
	IF span.status <> 0 THEN
		THIS^.AssertEquals_UDINT(TO_UDINT(E_StatusCode.STATUS_CODE_ERROR), TO_UDINT(span.status^.code), 'Expected an error code');
		THIS^.AssertTrue(span.status^.message <> 0, 'Expected a message');
		IF span.status^.message <> 0 THEN
			THIS^.AssertEquals_STRING('motor over temp', span.status^.message^.pString^, 'Expected the span to keep its own copy of the message');
		END_IF
	END_IF

	success := tracer.setSpanStatusError(pSpan:=ADR(emptySpan), message:='', failureReason=>reason);
	THIS^.AssertTrue(success, 'Expected an empty message to succeed');
	THIS^.AssertEquals_UDINT(TO_UDINT(E_TracerFailureReason.NA), TO_UDINT(reason), 'Expected no failure for an empty message');
	IF emptySpan.status <> 0 THEN
		THIS^.AssertEquals_UDINT(TO_UDINT(E_StatusCode.STATUS_CODE_ERROR), TO_UDINT(emptySpan.status^.code), 'Expected an error code without a message');
		THIS^.AssertTrue(emptySpan.status^.message = 0, 'Expected an empty message to leave no message');
	END_IF
	span.free();
	emptySpan.free();
TcUnit.TEST_FINISHED();
END_METHOD

(* The first status set wins: any later setSpanStatusOk or setSpanStatusError is refused
   with SPAN_STATUS_ALREADY_SET and leaves the status and its message unchanged. *)
METHOD testSetSpanStatusFirstWins : REFERENCE TO FB_Test
VAR
	resource: FB_Resource('');
	idGenerator: FB_MockIdGenerator;
	provider: FB_TracerProvider(resource:=resource, idGenerator:=idGenerator, sampler:=TcOtlp_GVL.defaultSampler);
	scope: FB_InstrumentationScope('tracer.test', '1.0.0', '');
	tracer: FB_Tracer(scope:=scope, provider:=provider);
	errorSpan: FB_Span;  // bare spans: the status setters need no identity
	okSpan: FB_Span;
	success: BOOL;
	reason: E_TracerFailureReason;
END_VAR
TcUnit.TEST('testSetSpanStatusFirstWins');
	tracer.setSpanStatusError(pSpan:=ADR(errorSpan), message:='first fault');

	success := tracer.setSpanStatusOk(pSpan:=ADR(errorSpan), failureReason=>reason);
	THIS^.AssertFalse(success, 'Expected OK after an error to be refused');
	THIS^.AssertEquals_UDINT(TO_UDINT(E_TracerFailureReason.SPAN_STATUS_ALREADY_SET), TO_UDINT(reason), 'Expected SPAN_STATUS_ALREADY_SET for OK after an error');

	success := tracer.setSpanStatusError(pSpan:=ADR(errorSpan), message:='second fault', failureReason=>reason);
	THIS^.AssertFalse(success, 'Expected a second error to be refused');
	THIS^.AssertEquals_UDINT(TO_UDINT(E_TracerFailureReason.SPAN_STATUS_ALREADY_SET), TO_UDINT(reason), 'Expected SPAN_STATUS_ALREADY_SET for a second error');

	THIS^.AssertTrue(errorSpan.status <> 0, 'Expected the first status to remain');
	IF errorSpan.status <> 0 THEN
		THIS^.AssertEquals_UDINT(TO_UDINT(E_StatusCode.STATUS_CODE_ERROR), TO_UDINT(errorSpan.status^.code), 'Expected the status to stay ERROR');
		THIS^.AssertTrue(errorSpan.status^.message <> 0, 'Expected the first message to remain');
		IF errorSpan.status^.message <> 0 THEN
			THIS^.AssertEquals_STRING('first fault', errorSpan.status^.message^.pString^, 'Expected the first message to win');
		END_IF
	END_IF

	tracer.setSpanStatusOk(pSpan:=ADR(okSpan));

	success := tracer.setSpanStatusError(pSpan:=ADR(okSpan), message:='late fault', failureReason=>reason);
	THIS^.AssertFalse(success, 'Expected an error after OK to be refused');
	THIS^.AssertEquals_UDINT(TO_UDINT(E_TracerFailureReason.SPAN_STATUS_ALREADY_SET), TO_UDINT(reason), 'Expected SPAN_STATUS_ALREADY_SET for an error after OK');

	success := tracer.setSpanStatusOk(pSpan:=ADR(okSpan), failureReason=>reason);
	THIS^.AssertFalse(success, 'Expected a second OK to be refused');
	THIS^.AssertEquals_UDINT(TO_UDINT(E_TracerFailureReason.SPAN_STATUS_ALREADY_SET), TO_UDINT(reason), 'Expected SPAN_STATUS_ALREADY_SET for a second OK');

	IF okSpan.status <> 0 THEN
		THIS^.AssertEquals_UDINT(TO_UDINT(E_StatusCode.STATUS_CODE_OK), TO_UDINT(okSpan.status^.code), 'Expected the status to stay OK');
		THIS^.AssertTrue(okSpan.status^.message = 0, 'Expected no message after the refused error');
	END_IF
	errorSpan.free();
	okSpan.free();
TcUnit.TEST_FINISHED();
END_METHOD

(* Writes distinct non-zero bytes into both identifiers. *)
METHOD _fillIds
VAR_IN_OUT
	traceId: FB_TraceId;
	spanId: FB_SpanId;
END_VAR
VAR
	_idx: UDINT;
	_bytes: ARRAY [0..15] OF BYTE;
END_VAR
FOR _idx := 0 TO SIZEOF(_bytes) - 1 DO
	_bytes[_idx] := TO_BYTE(_idx) + 1;
END_FOR
MEMCPY(ADR(traceId.bytes), ADR(_bytes), SIZEOF(traceId.bytes));

FOR _idx := 0 TO SIZEOF(_bytes) - 1 DO
	_bytes[_idx] := TO_BYTE(_idx) + 16#40;
END_FOR
MEMCPY(ADR(spanId.bytes), ADR(_bytes), SIZEOF(spanId.bytes));
END_METHOD

(* The context holds copies of the span's identifiers and trace state, so it stays intact
   after the span ends. *)
METHOD testGetSpanContextCopiesIdentity : REFERENCE TO FB_Test
VAR
	resource: FB_Resource('');
	idGenerator: FB_MockIdGenerator;
	provider: FB_TracerProvider(resource:=resource, idGenerator:=idGenerator, sampler:=TcOtlp_GVL.defaultSampler);
	scope: FB_InstrumentationScope('tracer.test', '1.0.0', '');
	tracer: FB_Tracer(scope:=scope, provider:=provider);
	pRemote: POINTER TO FB_SpanContext;
	pSpan: POINTER TO FB_Span;
	pContext: POINTER TO FB_SpanContext;
	traceId: FB_TraceId;
	spanId: FB_SpanId;
	pTraceState: POINTER TO FB_TraceState;
	traceStateText: T_MaxString := 'vendor=abc';
	success: BOOL;
	failureReason: E_TracerFailureReason;
END_VAR
TcUnit.TEST('testGetSpanContextCopiesIdentity');
	// a remote parent is the only way a span gets trace state; 16#301 is sampled, remoteness known, remote
	THIS^._fillIds(traceId:=traceId, spanId:=spanId);
	TraceStateFactory.parse(pDest:=pTraceState, pHeader:=ADR(traceStateText));
	ContextFactory.buildContext(
		pDest:=pRemote,
		pTraceId:=ADR(traceId),
		pSpanId:=ADR(spanId),
		pTraceState:=pTraceState,
		traceFlags:=16#301
	);
	IF pTraceState <> 0 THEN pTraceState^.delete(pSelf:=pTraceState); END_IF
	tracer.startSpan(name:='work').setParentUsingContext(pContext:=pRemote).build(pDest:=pSpan);
	IF pRemote <> 0 THEN pRemote^.delete(pSelf:=pRemote); END_IF
	THIS^.AssertTrue(pSpan <> 0 AND_THEN pSpan^.traceState <> 0, 'Expected the tracer to build a span with trace state');

	IF pSpan <> 0 AND_THEN pSpan^.traceState <> 0 THEN
		success := tracer.getSpanContext(pSpan:=pSpan, pDest:=pContext, failureReason=>failureReason);
		THIS^.AssertTrue(success, 'Expected getSpanContext to succeed for a span with an identity');
		THIS^.AssertEquals_UDINT(
			TO_UDINT(E_TracerFailureReason.NA),
			TO_UDINT(failureReason),
			'Expected no failure reason on success'
		);
		THIS^.AssertTrue(pContext <> 0, 'Expected getSpanContext to assign the destination');

		IF pContext <> 0 THEN
			THIS^.AssertTrue(pContext^.isValid(), 'Expected the context to be valid');
			THIS^.AssertTrue(
				MEMCMP(ADR(pContext^.traceId.bytes), ADR(pSpan^.traceId^.bytes), SIZEOF(pContext^.traceId.bytes)) = 0,
				'Expected the context to hold the span$'s trace id'
			);
			THIS^.AssertTrue(
				MEMCMP(ADR(pContext^.spanId.bytes), ADR(pSpan^.spanId^.bytes), SIZEOF(pContext^.spanId.bytes)) = 0,
				'Expected the context to hold the span$'s span id'
			);
			THIS^.AssertTrue(pContext^.traceState <> 0 AND_THEN pContext^.traceState <> pSpan^.traceState,
				'Expected the context to hold its own copy of the trace state');
			IF pContext^.traceState <> 0 THEN
				THIS^.AssertEquals_STRING('vendor=abc', pContext^.traceState^.pString^, 'Expected the trace state text to be copied');
			END_IF
		END_IF
	END_IF

	// the span is released first; the context must not depend on it
	IF pSpan <> 0 THEN pSpan^.delete(pSelf:=pSpan); END_IF
	IF pContext <> 0 AND_THEN pContext^.traceState <> 0 THEN
		THIS^.AssertEquals_STRING('vendor=abc', pContext^.traceState^.pString^, 'Expected the context$'s trace state to outlive the span');
	END_IF

	IF pContext <> 0 THEN pContext^.delete(pSelf:=pContext); END_IF
TcUnit.TEST_FINISHED();
END_METHOD

(* A context taken from a local span is known to be local: bit 8 is set and bit 9 is clear.
   A span without trace state gives a context without trace state. *)
METHOD testGetSpanContextIsLocal : REFERENCE TO FB_Test
VAR
	resource: FB_Resource('');
	idGenerator: FB_MockIdGenerator;
	provider: FB_TracerProvider(resource:=resource, idGenerator:=idGenerator, sampler:=TcOtlp_GVL.defaultSampler);
	scope: FB_InstrumentationScope('tracer.test', '1.0.0', '');
	tracer: FB_Tracer(scope:=scope, provider:=provider);
	pSpan: POINTER TO FB_Span;
	pContext: POINTER TO FB_SpanContext;
END_VAR
TcUnit.TEST('testGetSpanContextIsLocal');
	// a root span has no trace state
	tracer.startSpan(name:='work').build(pDest:=pSpan);
	THIS^.AssertTrue(pSpan <> 0, 'Expected the tracer to build a root span');

	IF pSpan <> 0 THEN
		tracer.getSpanContext(pSpan:=pSpan, pDest:=pContext);
		THIS^.AssertTrue(pContext <> 0, 'Expected getSpanContext to assign the destination');
		IF pContext <> 0 THEN
			THIS^.AssertFalse(pContext^.isRemote(), 'Expected a local span$'s context not to be remote');
			THIS^.AssertTrue(
				(pContext^.traceFlags AND TO_UDINT(E_SpanFlags.SPAN_FLAGS_CONTEXT_HAS_IS_REMOTE_MASK)) <> 0,
				'Expected remoteness to be marked as known'
			);
			THIS^.AssertTrue(
				(pContext^.traceFlags AND TO_UDINT(E_SpanFlags.SPAN_FLAGS_CONTEXT_IS_REMOTE_MASK)) = 0,
				'Expected the remote bit to be clear'
			);
			THIS^.AssertTrue(pContext^.traceState = 0, 'Expected no trace state when the span has none');
			pContext^.delete(pSelf:=pContext);
		END_IF
		pSpan^.delete(pSelf:=pSpan);
	END_IF
TcUnit.TEST_FINISHED();
END_METHOD

(* getSpanContext follows the VAR_IN_OUT pointer pattern: it never overwrites a context the
   caller already owns. *)
METHOD testGetSpanContextRejectsAssignedDestination : REFERENCE TO FB_Test
VAR
	resource: FB_Resource('');
	idGenerator: FB_MockIdGenerator;
	provider: FB_TracerProvider(resource:=resource, idGenerator:=idGenerator, sampler:=TcOtlp_GVL.defaultSampler);
	scope: FB_InstrumentationScope('tracer.test', '1.0.0', '');
	tracer: FB_Tracer(scope:=scope, provider:=provider);
	pSpan: POINTER TO FB_Span;
	pContext: POINTER TO FB_SpanContext;
	pFirst: POINTER TO FB_SpanContext;
	success: BOOL;
	reason: E_TracerFailureReason;
END_VAR
TcUnit.TEST('testGetSpanContextRejectsAssignedDestination');
	tracer.startSpan(name:='work').build(pDest:=pSpan);
	THIS^.AssertTrue(pSpan <> 0, 'Expected the tracer to build a root span');

	IF pSpan <> 0 THEN
		success := tracer.getSpanContext(pSpan:=pSpan, pDest:=pContext);
		THIS^.AssertTrue(success, 'Expected the first getSpanContext to succeed');
		pFirst := pContext;

		success := tracer.getSpanContext(pSpan:=pSpan, pDest:=pContext, failureReason=>reason);
		THIS^.AssertFalse(success, 'Expected getSpanContext into an assigned destination to fail');
		THIS^.AssertEquals_UDINT(TO_UDINT(E_TracerFailureReason.DESTINATION_ALREADY_ASSIGNED), TO_UDINT(reason), 'Expected DESTINATION_ALREADY_ASSIGNED');
		THIS^.AssertTrue(pContext = pFirst, 'Expected the destination pointer to be left alone');

		pSpan^.delete(pSelf:=pSpan);
	END_IF
	IF pContext <> 0 THEN pContext^.delete(pSelf:=pContext); END_IF
TcUnit.TEST_FINISHED();
END_METHOD

(* A span with no identity yet has nothing to snapshot, so getSpanContext refuses it with
   SPAN_INVALID and allocates nothing. *)
METHOD testGetSpanContextOnUnbuiltSpan : REFERENCE TO FB_Test
VAR
	resource: FB_Resource('');
	idGenerator: FB_MockIdGenerator;
	provider: FB_TracerProvider(resource:=resource, idGenerator:=idGenerator, sampler:=TcOtlp_GVL.defaultSampler);
	scope: FB_InstrumentationScope('tracer.test', '1.0.0', '');
	tracer: FB_Tracer(scope:=scope, provider:=provider);
	span: FB_Span;
	pContext: POINTER TO FB_SpanContext;
	success: BOOL;
	reason: E_TracerFailureReason;
END_VAR
TcUnit.TEST('testGetSpanContextOnUnbuiltSpan');
	success := tracer.getSpanContext(pSpan:=ADR(span), pDest:=pContext, failureReason=>reason);
	THIS^.AssertFalse(success, 'Expected getSpanContext to fail for a span without an identity');
	THIS^.AssertEquals_UDINT(TO_UDINT(E_TracerFailureReason.SPAN_INVALID), TO_UDINT(reason), 'Expected SPAN_INVALID');
	THIS^.AssertTrue(pContext = 0, 'Expected the destination to stay unassigned');
TcUnit.TEST_FINISHED();
END_METHOD

(* addSpanLink links a running span to a borrowed context, and pushSpanLink takes a link
   built with LinkFactory, clearing the caller's pointer. *)
METHOD testAddsLinksToRunningSpan : REFERENCE TO FB_Test
VAR
	resource: FB_Resource('');
	idGenerator: FB_MockIdGenerator;
	provider: FB_TracerProvider(resource:=resource, idGenerator:=idGenerator, sampler:=TcOtlp_GVL.defaultSampler);
	scope: FB_InstrumentationScope('tracer.test', '1.0.0', '');
	tracer: FB_Tracer(scope:=scope, provider:=provider);
	pTrigger: POINTER TO FB_Span;
	pSpan: POINTER TO FB_Span;
	pTriggerContext: POINTER TO FB_SpanContext;
	pLink: POINTER TO FB_Link;
	success: BOOL;
	reason: E_TracerFailureReason;
END_VAR
TcUnit.TEST('testAddsLinksToRunningSpan');
	tracer.startSpan(name:='trigger').build(pDest:=pTrigger);
	tracer.getSpanContext(pSpan:=pTrigger, pDest:=pTriggerContext);
	tracer.startSpan(name:='work').build(pDest:=pSpan);
	THIS^.AssertTrue(pSpan <> 0, 'Expected the span to build');

	success := tracer.addSpanLink(pSpan:=pSpan, pContext:=pTriggerContext, failureReason=>reason);
	THIS^.AssertTrue(success, 'Expected addSpanLink to succeed');
	THIS^.AssertEquals_UDINT(TO_UDINT(E_TracerFailureReason.NA), TO_UDINT(reason), 'Expected no failure from addSpanLink');
	// the context is borrowed, so the caller still owns it
	THIS^.AssertTrue(pTriggerContext <> 0, 'Expected the context to stay with the caller');

	LinkFactory.fromContext(pDest:=pLink, pContext:=pTriggerContext);
	success := tracer.pushSpanLink(pSpan:=pSpan, pLink:=pLink, failureReason=>reason);
	THIS^.AssertTrue(success, 'Expected pushSpanLink to succeed');
	THIS^.AssertTrue(pLink = 0, 'Expected pushSpanLink to take the link');

	success := tracer.addSpanLink(pSpan:=pSpan, pContext:=0, failureReason=>reason);
	THIS^.AssertFalse(success, 'Expected addSpanLink to refuse a null context');
	THIS^.AssertEquals_UDINT(TO_UDINT(E_TracerFailureReason.LINK_CONTEXT_POINTER_NULL), TO_UDINT(reason), 'Expected LINK_CONTEXT_POINTER_NULL');

	success := tracer.pushSpanLink(pSpan:=pSpan, pLink:=pLink, failureReason=>reason);
	THIS^.AssertFalse(success, 'Expected pushSpanLink to refuse a null link');
	THIS^.AssertEquals_UDINT(TO_UDINT(E_TracerFailureReason.LINK_POINTER_NULL), TO_UDINT(reason), 'Expected LINK_POINTER_NULL');

	IF pSpan <> 0 THEN
		THIS^.AssertEquals_UDINT(2, pSpan^.links.count, 'Expected two links on the running span');
	END_IF
	IF pTriggerContext <> 0 THEN pTriggerContext^.delete(pSelf:=pTriggerContext); END_IF
	tracer.discardSpan(pSpan:=pSpan);
	tracer.discardSpan(pSpan:=pTrigger);
TcUnit.TEST_FINISHED();
END_METHOD

(* Attributes set on a running span are owned by the span. *)
METHOD testSetsRunningSpanAttributes : REFERENCE TO FB_Test
VAR
	resource: FB_Resource('');
	idGenerator: FB_MockIdGenerator;
	provider: FB_TracerProvider(resource:=resource, idGenerator:=idGenerator, sampler:=TcOtlp_GVL.defaultSampler);
	scope: FB_InstrumentationScope('tracer.test', '1.0.0', '');
	tracer: FB_Tracer(scope:=scope, provider:=provider);
	pSpan: POINTER TO FB_Span;
	setpoint: DINT := 42;
	success: BOOL;
	reason: E_TracerFailureReason;
END_VAR
TcUnit.TEST('testSetsRunningSpanAttributes');
	tracer.startSpan(name:='span').build(pDest:=pSpan);
	THIS^.AssertTrue(pSpan <> 0, 'Expected the span to build');

	success := tracer.setSpanStringAttribute(pSpan:=pSpan, key:='skid', value:='A', failureReason=>reason);
	THIS^.AssertTrue(success, 'Expected setSpanStringAttribute to succeed');
	THIS^.AssertEquals_UDINT(TO_UDINT(E_TracerFailureReason.NA), TO_UDINT(reason), 'Expected no failure from setSpanStringAttribute');

	success := tracer.setSpanNumberAttribute(pSpan:=pSpan, key:='setpoint', value:=setpoint, failureReason=>reason);
	THIS^.AssertTrue(success, 'Expected setSpanNumberAttribute to succeed');
	THIS^.AssertEquals_UDINT(TO_UDINT(E_TracerFailureReason.NA), TO_UDINT(reason), 'Expected no failure from setSpanNumberAttribute');

	IF pSpan <> 0 THEN
		THIS^.AssertEquals_UDINT(2, pSpan^.attributes.count, 'Expected both attributes on the span');
	END_IF
	tracer.discardSpan(pSpan:=pSpan);
TcUnit.TEST_FINISHED();
END_METHOD

(* discardSpan releases a running span without handing it to the provider, and clears the
   caller's pointer. *)
METHOD testDiscardSpanReleasesSpan : REFERENCE TO FB_Test
VAR
	resource: FB_Resource('');
	idGenerator: FB_MockIdGenerator;
	provider: FB_TracerProvider_ForInspection(resource:=resource, idGenerator:=idGenerator, sampler:=TcOtlp_GVL.defaultSampler);
	scope: FB_InstrumentationScope('tracer.test', '1.0.0', '');
	tracer: FB_Tracer(scope:=scope, provider:=provider);
	pSpan: POINTER TO FB_Span;
	success: BOOL;
	reason: E_TracerFailureReason;
END_VAR
TcUnit.TEST('testDiscardSpanReleasesSpan');
	tracer.startSpan(name:='abandoned').build(pDest:=pSpan);
	THIS^.AssertTrue(pSpan <> 0, 'Expected the span to build');

	success := tracer.discardSpan(pSpan:=pSpan, failureReason=>reason);
	THIS^.AssertTrue(success, 'Expected discardSpan to succeed');
	THIS^.AssertEquals_UDINT(TO_UDINT(E_TracerFailureReason.NA), TO_UDINT(reason), 'Expected no failure');
	THIS^.AssertTrue(pSpan = 0, 'Expected the caller$'s pointer to be cleared');
	THIS^.AssertEquals_UDINT(0, provider.spans.count, 'Expected nothing to be queued');
TcUnit.TEST_FINISHED();
END_METHOD

(* Every method for a running span refuses a null span with SPAN_POINTER_NULL, so callers need
   no null check of their own. pushSpanLink still releases the link it was given. *)
METHOD testRunningSpanMethodsRejectNullSpan : REFERENCE TO FB_Test
VAR
	resource: FB_Resource('');
	idGenerator: FB_MockIdGenerator;
	provider: FB_TracerProvider(resource:=resource, idGenerator:=idGenerator, sampler:=TcOtlp_GVL.defaultSampler);
	scope: FB_InstrumentationScope('tracer.test', '1.0.0', '');
	tracer: FB_Tracer(scope:=scope, provider:=provider);
	pSpan: POINTER TO FB_Span;
	pRoot: POINTER TO FB_Span;
	pContext: POINTER TO FB_SpanContext;
	pLink: POINTER TO FB_Link;
	setpoint: DINT := 42;
	success: BOOL;
	reason: E_TracerFailureReason;
END_VAR
TcUnit.TEST('testRunningSpanMethodsRejectNullSpan');
	success := tracer.setSpanStatusOk(pSpan:=pSpan, failureReason=>reason);
	THIS^.AssertFalse(success, 'Expected setSpanStatusOk to refuse a null span');
	THIS^.AssertEquals_UDINT(TO_UDINT(E_TracerFailureReason.SPAN_POINTER_NULL), TO_UDINT(reason), 'Expected SPAN_POINTER_NULL from setSpanStatusOk');

	success := tracer.setSpanStatusError(pSpan:=pSpan, message:='boom', failureReason=>reason);
	THIS^.AssertFalse(success, 'Expected setSpanStatusError to refuse a null span');
	THIS^.AssertEquals_UDINT(TO_UDINT(E_TracerFailureReason.SPAN_POINTER_NULL), TO_UDINT(reason), 'Expected SPAN_POINTER_NULL from setSpanStatusError');

	success := tracer.getSpanContext(pSpan:=pSpan, pDest:=pContext, failureReason=>reason);
	THIS^.AssertFalse(success, 'Expected getSpanContext to refuse a null span');
	THIS^.AssertEquals_UDINT(TO_UDINT(E_TracerFailureReason.SPAN_POINTER_NULL), TO_UDINT(reason), 'Expected SPAN_POINTER_NULL from getSpanContext');
	THIS^.AssertTrue(pContext = 0, 'Expected getSpanContext to allocate nothing');

	success := tracer.setSpanStringAttribute(pSpan:=pSpan, key:='k', value:='v', failureReason=>reason);
	THIS^.AssertFalse(success, 'Expected setSpanStringAttribute to refuse a null span');
	THIS^.AssertEquals_UDINT(TO_UDINT(E_TracerFailureReason.SPAN_POINTER_NULL), TO_UDINT(reason), 'Expected SPAN_POINTER_NULL from setSpanStringAttribute');

	success := tracer.setSpanNumberAttribute(pSpan:=pSpan, key:='k', value:=setpoint, failureReason=>reason);
	THIS^.AssertFalse(success, 'Expected setSpanNumberAttribute to refuse a null span');
	THIS^.AssertEquals_UDINT(TO_UDINT(E_TracerFailureReason.SPAN_POINTER_NULL), TO_UDINT(reason), 'Expected SPAN_POINTER_NULL from setSpanNumberAttribute');

	// a real context and link, so the null span is the only thing wrong
	tracer.startSpan(name:='root').build(pDest:=pRoot);
	tracer.getSpanContext(pSpan:=pRoot, pDest:=pContext);

	success := tracer.addSpanLink(pSpan:=pSpan, pContext:=pContext, failureReason=>reason);
	THIS^.AssertFalse(success, 'Expected addSpanLink to refuse a null span');
	THIS^.AssertEquals_UDINT(TO_UDINT(E_TracerFailureReason.SPAN_POINTER_NULL), TO_UDINT(reason), 'Expected SPAN_POINTER_NULL from addSpanLink');

	LinkFactory.fromContext(pDest:=pLink, pContext:=pContext);
	THIS^.AssertTrue(pLink <> 0, 'Expected a link to push');
	success := tracer.pushSpanLink(pSpan:=pSpan, pLink:=pLink, failureReason=>reason);
	THIS^.AssertFalse(success, 'Expected pushSpanLink to refuse a null span');
	THIS^.AssertEquals_UDINT(TO_UDINT(E_TracerFailureReason.SPAN_POINTER_NULL), TO_UDINT(reason), 'Expected SPAN_POINTER_NULL from pushSpanLink');
	THIS^.AssertTrue(pLink = 0, 'Expected pushSpanLink to release the refused link');

	success := tracer.discardSpan(pSpan:=pSpan, failureReason=>reason);
	THIS^.AssertFalse(success, 'Expected discardSpan to refuse a null span');
	THIS^.AssertEquals_UDINT(TO_UDINT(E_TracerFailureReason.SPAN_POINTER_NULL), TO_UDINT(reason), 'Expected SPAN_POINTER_NULL from discardSpan');

	IF pContext <> 0 THEN pContext^.delete(pSelf:=pContext); END_IF
	tracer.discardSpan(pSpan:=pRoot);
TcUnit.TEST_FINISHED();
END_METHOD

(* addLink links the span to other contexts, in the order they are added, without making it
   a child. The contexts are borrowed. *)
METHOD testAddsLinks : REFERENCE TO FB_Test
VAR
	resource: FB_Resource('');
	idGenerator: FB_MockIdGenerator;
	provider: FB_TracerProvider(resource:=resource, idGenerator:=idGenerator, sampler:=TcOtlp_GVL.defaultSampler);
	scope: FB_InstrumentationScope('tracer.test', '1.0.0', '');
	tracer: FB_Tracer(scope:=scope, provider:=provider);
	pTrigger: POINTER TO FB_Span;
	pSpan: POINTER TO FB_Span;
	pTriggerContext: POINTER TO FB_SpanContext;
	pRemote: POINTER TO FB_SpanContext;
	pLink: POINTER TO FB_Link;
	traceId: FB_TraceId;
	spanId: FB_SpanId;
	success: BOOL;
	reason: E_TracerFailureReason;
END_VAR
TcUnit.TEST('testAddsLinks');
	tracer.startSpan(name:='trigger').build(pDest:=pTrigger);
	IF pTrigger <> 0 THEN tracer.getSpanContext(pSpan:=pTrigger, pDest:=pTriggerContext); END_IF
	MEMSET(ADR(traceId.bytes), 16#AA, SIZEOF(traceId.bytes));
	MEMSET(ADR(spanId.bytes), 16#BB, SIZEOF(spanId.bytes));
	ContextFactory.buildContext(pDest:=pRemote, pTraceId:=ADR(traceId), pSpanId:=ADR(spanId), pTraceState:=0, traceFlags:=16#301);

	success := tracer
		.startSpan(name:='work')
		.addLink(pContext:=pTriggerContext)
		.addLink(pContext:=pRemote)
		.build(pDest:=pSpan, failureReason=>reason);
	THIS^.AssertTrue(success, 'Expected a span with links to build');
	THIS^.AssertEquals_UDINT(TO_UDINT(E_TracerFailureReason.NA), TO_UDINT(reason), 'Expected no failure reason');

	// the contexts are borrowed, so they can be released before the span
	IF pTriggerContext <> 0 THEN pTriggerContext^.delete(pSelf:=pTriggerContext); END_IF
	IF pRemote <> 0 THEN pRemote^.delete(pSelf:=pRemote); END_IF

